RoboDK station: verify_station_copy.rdk

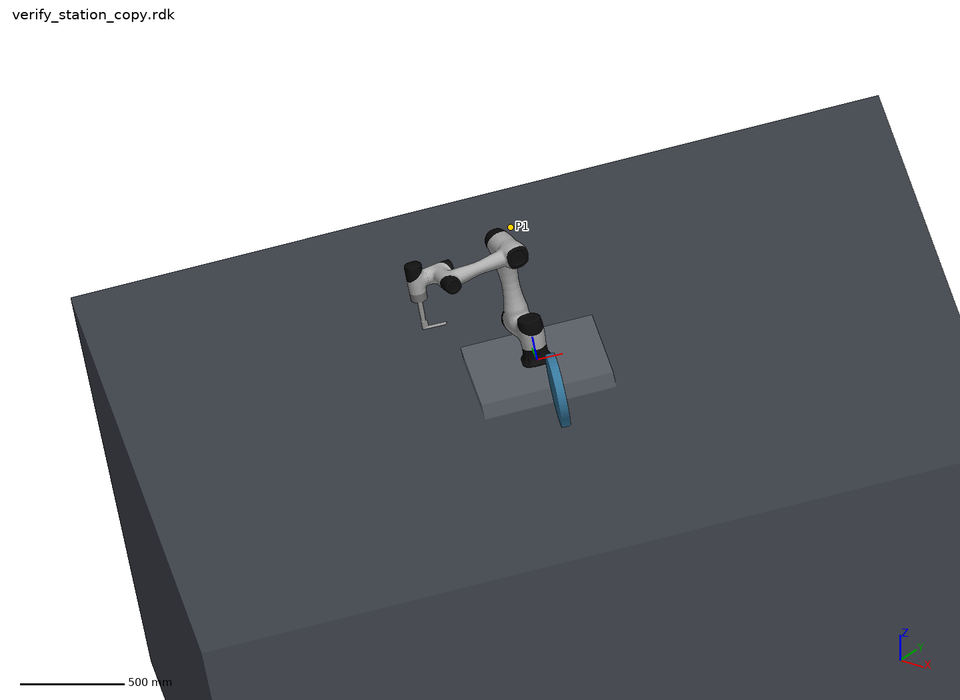
[picture v0: the station drawn from its stored meshes, robots at their saved joint values, targets as dots, program paths as lines]
Station 新建工作站 (1) (saved by RoboDK 5.9.0). Poses are relative to the parent item; angles as X-Y-Z fixed-axis rotations.
Station parameters (name, value as stored): Trace_Render_Style, 0
  - Python program TCP真实运动_升级前备份_20260910_170410 (listed below)
  - Python program 方向角计算 (listed below)
  - frame Dobot CR5 Base at (213.88, 904.45, 25.18) mm, rotated rx -0.42 ry -9.85 rz 44.17 deg
    - robot Dobot CR5: 6 axes, payload 5 kg, reach 900 mm, repeatability 0.03 mm, weight 23 kg
        modified DH rows (alpha deg, a mm, theta deg, d mm): 0, 0, 0, 147; 90, 0, 90, 0; 0, 427, 0, 0; 0, 357, -90, 141; -90, 0, 0, 116; 90, 0, 180, 100.5
        joint limits [-360, -360, -160, -360, -360, -360] to [360, 360, 160, 360, 360, 360]; home [0, 0, -90, 90, 90, 0]; saved at [-163.62, -0.936, -91.282, 2.218, 90, 106.38]
      - tool , TCP at (0, 0, 159.63) mm, size 120.1 x 159.6 x 24.6 mm, geometry from bs1.stp
    - target P1 (joint target) at (-20.1, -241.48, 846.75) mm, rotated rx -90 ry 1.35 rz 179.96 deg; joints [0, -37.451, 84.112, -46.661, 0, 0] of Dobot CR5
    - object  at (0, 0, 0) mm, rotated rx 0 ry -1.35 rz -0.05 deg, size 650 x 650 x 80 mm
    - object  at (0, 0, 0) mm, rotated rx 0 ry -1.35 rz -0.05 deg, size 4000 x 4000 x 2000 mm
    - object  at (0, -956, 300) mm, rotated rx 139.77 ry 89.72 rz -40.3 deg, size 360 x 360 x 40 mm
  - Python program TCP仿真_升级前备份_20260909_173616 (listed below)
  - Python program TCP仿真_升级前备份_20260910_161757 (listed below)
  - Python program TCP仿真_升级前备份_20260910_164419 (listed below)
  - Python program test (listed below)
  - Python program 机械臂法兰真实运动 (listed below)
  - Python program TCP真实运动_到位复核前备份_20260910_172919 (listed below)
  - Python program TCP真实运动 (listed below)
  - Python program TCP仿真_退让换向升级前 (listed below)
  - Python program TCP仿真 (listed below)
  - Python program 机械臂TCP仿真_副本 (listed below)

--- Python program TCP真实运动_升级前备份_20260910_170410 ---
# -*- coding: utf-8 -*-
"""
RoboDK 实机运动控制（基于 robodk_movej_diag.py 的成功模式）
- 单点：TCP 输入 -> IK 检测 -> MoveL/MoveJ 执行
- 连续轨迹：坐标列表 -> 逐点 IK 检测 -> MoveJ+MoveL 序列
模式：RUNMODE_RUN_ROBOT + robot.Connect()
"""

from robodk.robolink import *
from robodk.robomath import *
import tkinter as tk
from tkinter import ttk, scrolledtext, filedialog
import time
import math
import json

ROBOT_SPEED = 20.0
NL = chr(10)

RDK = Robolink()

def fanuc_to_pose(x, y, z, rx, ry, rz):
    return Fanuc_2_Pose([x, y, z, rx, ry, rz])

def pose_to_fanuc(pose):
    return Pose_2_Fanuc(pose)

# ---- 获取机器人 ----
robot = RDK.Item('', ITEM_TYPE_ROBOT)
if not robot.Valid():
    raise Exception("未找到机器人")

# ---- 全局变量 ----
text_points = None
text_log = None
record_text = None
entries_single = None
entries_joint = None
move_type = None
trajectory_records = []
_connected = False

# ============================================================
# 日志
# ============================================================
def log(s):
    print(s)
    if text_log:
        text_log.insert(tk.END, str(s) + NL)
        text_log.see(tk.END)
        root.update_idletasks()

# ============================================================
# 连接（只连一次，复用）
# ============================================================
def ensure_connected():
    global _connected
    if _connected:
        return True
    try:
        robot.Connect()
        time.sleep(1.5)
        status, msg = robot.ConnectedState()
        log("连接状态: %s, %s" % (status, msg))
        RDK.setRunMode(RUNMODE_RUN_ROBOT)
        log("RunMode: %s" % RDK.RunMode())
        if status < 0:
            _connected = False
            log("机器人连接未建立，状态=%s：%s" % (status, msg))
            return False
        _connected = True
        return True
    except Exception as e:
        log("连接失败: %s" % e)
        return False

# ============================================================
# 解析坐标
# ============================================================
def parse_points():
    if not text_points:
        return []
    raw = text_points.get("1.0", tk.END)
    points = []
    for line in raw.strip().split(NL):
        line = line.strip()
        if not line or line.startswith("#"):
            continue
        try:
            vals = [float(v.strip()) for v in line.split(",")]
            if len(vals) >= 6:
                points.append(vals[:6])
        except ValueError:
            pass
    return points

# ============================================================
# 读取当前位置
# ============================================================
def read_current(entries=None):
    try:
        pose = robot.Pose()
        v = pose_to_fanuc(pose)
        log("")
        log("当前 TCP：X=%.3f Y=%.3f Z=%.3f Rx=%.3f Ry=%.3f Rz=%.3f" % tuple(v[:6]))
    except Exception as e:
        log("读取失败：%s" % e)

def fill_current(entries=None):
    try:
        pose = robot.Pose()
        v = pose_to_fanuc(pose)
        if entries:
            for e, val in zip(entries, v):
                e.delete(0, tk.END)
                e.insert(0, "%.3f" % val)
        log("当前 TCP 已填入")
    except Exception as e:
        log("读取失败：%s" % e)

# ============================================================
# IK 检测
# 注意：SolveIK 显式使用当前 Tool + Reference，和 MoveL/MoveJ 保持一致。
# ============================================================
def check_ik_single(entries=None):
    if not entries:
        return
    try:
        values = [float(e.get()) for e in entries]
    except ValueError:
        log("输入无效")
        return

    x, y, z, rx, ry, rz = values
    target = fanuc_to_pose(x, y, z, rx, ry, rz)
    log("")
    log("目标：X=%.3f Y=%.3f Z=%.3f Rx=%.3f Ry=%.3f Rz=%.3f" % (x, y, z, rx, ry, rz))

    try:
        tool_pose = robot.PoseTool()
        frame_pose = robot.PoseFrame()
        joints = robot.SolveIK(target, tool=tool_pose, reference=frame_pose)
        if joints is None:
            log("IK 不可达")
        else:
            q = joints.list()
            if len(q) < 6:
                log("IK 返回关节数量异常：%d，原始数据=%r" % (len(q), q))
                return
            log("IK 可达")
            log("  关节：J1=%.2f J2=%.2f J3=%.2f J4=%.2f J5=%.2f J6=%.2f" % tuple(q[:6]))
    except Exception as e:
        log("检测失败：%s" % e)

def check_all_ik():
    points = parse_points()
    if not points:
        log("没有有效点")
        return

    log("")
    log("========== 检测全部 %d 个点 ==========" % len(points))
    all_ok = True
    for i, p in enumerate(points):
        try:
            target = fanuc_to_pose(*p)
            joints = robot.SolveIK(target, tool=robot.PoseTool(), reference=robot.PoseFrame())
            if joints is None:
                log("  P%d: 不可达" % (i+1))
                all_ok = False
            else:
                q = joints.list()
                if len(q) < 6:
                    raise ValueError("IK 返回关节数量异常: %d, raw=%r" % (len(q), q))
                log("  P%d: 可达  J1=%.1f J2=%.1f J3=%.1f J4=%.1f J5=%.1f J6=%.1f" % (i+1, *q[:6]))
        except Exception as e:
            log("  P%d: 检测失败 %s" % (i+1, e))
            all_ok = False
    if all_ok:
        log("全部 %d 个点可达" % len(points))
    else:
        log("存在不可达点，执行时会跳过")

# ============================================================
# 执行单点
# ============================================================
def execute_single(entries=None, mtype="MoveL"):
    if not entries:
        return
    try:
        values = [float(e.get()) for e in entries]
    except ValueError:
        log("输入无效")
        return

    x, y, z, rx, ry, rz = values
    target = fanuc_to_pose(x, y, z, rx, ry, rz)
    log("")
    log("目标：X=%.3f Y=%.3f Z=%.3f Rx=%.3f Ry=%.3f Rz=%.3f" % (x, y, z, rx, ry, rz))

    try:
        tool_pose = robot.PoseTool()
        frame_pose = robot.PoseFrame()
        joints = robot.SolveIK(target, tool=tool_pose, reference=frame_pose)
        if joints is None:
            log("IK 不可达，取消执行")
            return
        q = joints.list()
        if len(q) < 6:
            log("IK 返回关节数量异常：%d，取消执行；原始数据=%r" % (len(q), q))
            return
        log("IK 可达：J1=%.2f J2=%.2f J3=%.2f J4=%.2f J5=%.2f J6=%.2f" % tuple(q[:6]))
    except Exception as e:
        log("IK 检查失败：%s" % e)
        return

    if not ensure_connected():
        return

    try:
        robot.setPoseFrame(robot.PoseFrame())
        robot.setPoseTool(robot.PoseTool())
        robot.setSpeed(ROBOT_SPEED)
        log("发送 %s..." % mtype)
        if mtype == "MoveJ":
            robot.MoveJ(target)
        else:
            robot.MoveL(target)
        log("执行完成")
    except Exception as e:
        log("失败: %s: %s" % (type(e).__name__, e))

# ============================================================
# 连续运动：选项卡3直接输入 TCP / 关节点，逐点检查后加入轨迹
# ============================================================
trajectory_records = []
record_text = None
traj_entries = None
traj_type = None
singular_var = None
j6_direction_var = None


def _parse_six_from_entries(entries, label):
    if not entries or len(entries) != 6:
        log("%s输入框异常：需要 6 个值" % label)
        return None
    try:
        vals = [float(e.get().strip()) for e in entries]
    except (ValueError, AttributeError):
        log("%s输入无效：6 个值必须全部为数字" % label)
        return None
    if not all(math.isfinite(v) for v in vals):
        log("%s输入无效：不能包含 NaN 或无穷值" % label)
        return None
    return vals


def _check_tcp_reachable(vals):
    """检查单个 TCP 点 IK 是否可达，返回 (True, target, joints)。"""
    try:
        target = fanuc_to_pose(*vals)
        tool_pose = robot.PoseTool()
        frame_pose = robot.PoseFrame()
        joints = robot.SolveIK(target, tool=tool_pose, reference=frame_pose)

        if joints is None:
            log("TCP IK：不可达")
            return False, None, None

        q = joints.list()
        if len(q) < 6:
            log("TCP IK：返回关节数量异常：%r" % q)
            return False, None, None

        log("TCP IK：可达")
        log("  IK关节：J1=%.2f J2=%.2f J3=%.2f J4=%.2f J5=%.2f J6=%.2f" % tuple(q[:6]))
        return True, target, q[:6]
    except Exception as e:
        log("TCP IK 检查失败：%s: %s" % (type(e).__name__, e))
        return False, None, None


def _check_tcp_segment_continuous(prev_vals, curr_vals, segment_index, samples=20):
    """检查前一个 TCP 点到当前 TCP 点之间的整段插补路径 IK 连续可达性。

    暂不考虑障碍物，只对 TCP 位姿做线性插值，并对每个采样位姿执行 SolveIK。
    起点和终点也包含在采样检查中。
    """
    if prev_vals is None:
        return True

    log("开始检查 P%d -> P%d 的 TCP 连续 IK（%d 个采样点）" %
        (segment_index - 1, segment_index, samples + 1))

    tool_pose = robot.PoseTool()
    frame_pose = robot.PoseFrame()

    for k in range(samples + 1):
        t = float(k) / float(samples)
        vals = [prev_vals[i] + (curr_vals[i] - prev_vals[i]) * t for i in range(6)]
        try:
            pose = fanuc_to_pose(*vals)
            joints = robot.SolveIK(pose, tool=tool_pose, reference=frame_pose)
            if joints is None:
                log("  P%d -> P%d：第 %d/%d 个采样点 IK 不可达，t=%.3f" %
                    (segment_index - 1, segment_index, k + 1, samples + 1, t))
                log("  TCP：X=%.3f Y=%.3f Z=%.3f Rx=%.3f Ry=%.3f Rz=%.3f" % tuple(vals))
                return False
            q = joints.list()
            if len(q) < 6:
                log("  P%d -> P%d：第 %d 个采样点 IK 返回异常：%r" %
                    (segment_index - 1, segment_index, k + 1, q))
                return False
        except Exception as e:
            log("  P%d -> P%d：第 %d 个采样点 IK 检查失败：%s: %s" %
                (segment_index - 1, segment_index, k + 1, type(e).__name__, e))
            return False

    log("P%d -> P%d：连续 IK 检查通过" % (segment_index - 1, segment_index))
    return True


def _check_joint_reachable(q):
    """兼容旧代码：关节点不做可达性/限位检查，输入合法即可加入。"""
    return True


def refresh_record_list():
    if record_text is None:
        return

    record_text.delete("1.0", tk.END)

    for i, rec in enumerate(trajectory_records, 1):
        kind = rec["type"]
        vals = rec["values"]

        if kind == "TCP":
            mark = " [J6特异点 %s180°]" % ("+" if rec.get("j6_delta", 180) >= 0 else "-") if rec.get("singular", False) else ""
            record_text.insert(
                tk.END,
                "P%-3d [TCP]%s   X=%9.3f Y=%9.3f Z=%9.3f Rx=%8.3f Ry=%8.3f Rz=%8.3f%s" %
                (i, mark, *vals, NL)
            )
        else:
            record_text.insert(
                tk.END,
                "P%-3d [JNT]   J1=%8.3f J2=%8.3f J3=%8.3f J4=%8.3f J5=%8.3f J6=%8.3f%s" %
                (i, *vals, NL)
            )


def add_and_check_trajectory_point():
    """
    选项卡3逐点输入：
    - 普通 TCP：立即做端点 IK，并检查与前一个普通 TCP 点之间的连续 IK。
    - TCP 末端特异点：跳过 IK；要求与前一个普通 TCP 点 XYZ 相同，执行时仅 J6 转 ±180°。
    - 关节：不做 IK/限位检查，只将角度规范到 (-180°, 180°]。
    注意：这些检查只在“加入点”时完成；正式实机执行时不再做轨迹预检。
    """
    kind = traj_type.get()
    vals = _parse_six_from_entries(traj_entries, kind)
    if vals is None:
        return

    log("")
    log("========== 检查连续运动第 %d 点 ==========" % (len(trajectory_records) + 1))

    is_singular = bool(singular_var.get()) if (kind == "TCP" and singular_var is not None) else False
    j6_delta = int(j6_direction_var.get()) if (j6_direction_var is not None) else 180

    if kind == "TCP" and is_singular:
        if not trajectory_records:
            log("末端特异点不能作为第一个点：需要先有一个起始运动点。")
            return
        prev = trajectory_records[-1]
        if prev["type"] != "TCP" or prev.get("singular", False):
            log("末端特异点前一项必须是普通 TCP 点。")
            return
        prev_vals = prev["values"]
        pos_err = math.sqrt(sum((vals[k] - prev_vals[k]) ** 2 for k in range(3)))
        if pos_err > 1e-3:
            log("末端特异点未加入：XYZ 必须与前一个普通 TCP 点相同。")
            log("  与前一点位置差：%.6f mm" % pos_err)
            return
        try:
            target = fanuc_to_pose(*vals)
        except Exception as e:
            log("末端特异点姿态转换失败：%s: %s" % (type(e).__name__, e))
            return

        trajectory_records.append({
            "type": "TCP", "values": vals[:], "target": target, "joints": None,
            "singular": True, "j6_delta": j6_delta,
        })
        log("P%d [TCP-特异点]：已加入，跳过 IK。" % len(trajectory_records))
        log("  执行时保持 J1~J5 不变，仅让 J6 转 %+d°。" % j6_delta)
        if singular_var is not None:
            singular_var.set(False)
        refresh_record_list()
        return

    if kind == "TCP":
        ok, target, joints = _check_tcp_reachable(vals)
        if not ok:
            log("该 TCP 点未加入轨迹。")
            return

        # 只在点加入阶段检查连续 IK；实机正式执行时不再重复预检。
        if trajectory_records and trajectory_records[-1]["type"] == "TCP" and not trajectory_records[-1].get("singular", False):
            prev_vals = trajectory_records[-1]["values"]
            segment_no = len(trajectory_records) + 1
            if not _check_tcp_segment_continuous(prev_vals, vals, segment_no, samples=20):
                log("P%d [TCP]：上一普通 TCP 点到当前点的连续 IK 检查失败，该点未加入轨迹。" % segment_no)
                return

        trajectory_records.append({
            "type": "TCP", "values": vals[:], "target": target, "joints": joints,
            "singular": False, "j6_delta": 0,
        })
        log("P%d [TCP]：检查通过，已加入连续运动。" % len(trajectory_records))
    else:
        corrected = []
        for v in vals:
            v = ((v + 180.0) % 360.0) - 180.0
            if v <= -180.0:
                v = 180.0
            corrected.append(v)
        if corrected != vals:
            log("关节点角度已自动纠正到 (-180°, 180°]：")
            log("  原始：" + "  ".join("J%d=%+.3f°" % (i + 1, vals[i]) for i in range(6)))
            log("  修正：" + "  ".join("J%d=%+.3f°" % (i + 1, corrected[i]) for i in range(6)))
        trajectory_records.append({
            "type": "JOINT", "values": corrected[:], "target": None, "joints": corrected[:],
            "singular": False, "j6_delta": 0,
        })
        log("P%d [JNT]：未做 IK 检查，角度规范化后已加入连续运动。" % len(trajectory_records))

    refresh_record_list()


def _write_values_to_traj_entries(values, label):
    if not traj_entries or len(traj_entries) != 6:
        log("连续运动输入框异常：无法写入当前%s" % label)
        return False
    for e, val in zip(traj_entries, values[:6]):
        e.delete(0, tk.END)
        e.insert(0, "%.3f" % float(val))
    log("当前%s已写入选项卡3输入框" % label)
    return True


def read_current_tcp_to_traj():
    """读取当前 RoboDK TCP，并写入选项卡3的 TCP 输入框。"""
    try:
        pose = robot.Pose()
        vals = pose_to_fanuc(pose)
        log("========== 读取当前 TCP -> 选项卡3 ==========")
        log("X=%+.3f Y=%+.3f Z=%+.3f Rx=%+.3f Ry=%+.3f Rz=%+.3f" % tuple(vals))
        if traj_type.get() != "TCP":
            traj_type.set("TCP")
            _update_traj_labels_and_defaults()
        return _write_values_to_traj_entries(vals, "TCP")
    except Exception as e:
        log("读取当前 TCP 失败：%s: %s" % (type(e).__name__, e))
        return False


def read_current_joints_to_traj():
    """读取 RoboDK Robot Item 当前关节，并写入选项卡3的关节输入框。"""
    q = read_current_joints(None)
    if q is None or len(q) < 6:
        return False
    log("========== 读取当前关节 -> 选项卡3 ==========")
    if traj_type.get() != "JOINT":
        traj_type.set("JOINT")
        _update_traj_labels_and_defaults()
    return _write_values_to_traj_entries(q, "关节")


def clear_trajectory_input():
    if not traj_entries:
        return

    for e in traj_entries:
        e.delete(0, tk.END)

    if traj_type.get() == "TCP":
        defaults = ["0.000", "-241.500", "1047.000", "-90.000", "0.000", "180.000"]
    else:
        defaults = ["0.000"] * 6

    for e, val in zip(traj_entries, defaults):
        e.insert(0, val)




def import_trajectory():
    """
    从仿真程序导出的 JSON 轨迹文件导入到实机连续运动列表。

    重要：这里不做连续轨迹预检，不做 MoveJ TCP 轨迹预检。
    普通 TCP 如果 JSON 中没有保存 IK 关节，则只针对该点单独 SolveIK，
    用于得到实机执行所需的目标关节；这不是连续轨迹预检。
    """
    filepath = filedialog.askopenfilename(
        title="导入仿真轨迹",
        defaultextension=".json",
        filetypes=[("JSON 轨迹文件", "*.json"), ("所有文件", "*.*")]
    )
    if not filepath:
        return

    try:
        with open(filepath, "r", encoding="utf-8") as f:
            data = json.load(f)

        if not isinstance(data, list):
            raise ValueError("轨迹文件顶层必须是列表。")

        imported = []
        for idx, item in enumerate(data, 1):
            if not isinstance(item, dict):
                raise ValueError("P%d 不是对象格式。" % idx)

            kind = str(item.get("type", "")).upper()
            if kind == "JNT":
                kind = "JOINT"
            if kind not in ("TCP", "JOINT"):
                raise ValueError("P%d type 不支持：%r" % (idx, item.get("type")))

            values = item.get("values")
            if not isinstance(values, list) or len(values) != 6:
                raise ValueError("P%d values 必须是长度为6的列表。" % idx)
            try:
                values = [float(v) for v in values]
            except (TypeError, ValueError):
                raise ValueError("P%d values 必须全部为数字。" % idx)
            if not all(math.isfinite(v) for v in values):
                raise ValueError("P%d values 不能包含 NaN 或无穷值。" % idx)

            is_singular = bool(item.get("singular", False)) and kind == "TCP"
            j6_delta = int(item.get("j6_delta", 180)) if is_singular else 0
            if is_singular and j6_delta not in (-180, 180):
                raise ValueError("P%d 特异点 j6_delta 只能是 +180 或 -180。" % idx)

            if kind == "JOINT":
                # 与手动输入保持一致：自动规范到 (-180,180]。
                corrected = []
                for v in values:
                    v = ((v + 180.0) % 360.0) - 180.0
                    if v <= -180.0:
                        v = 180.0
                    corrected.append(v)
                values = corrected
                imported.append({
                    "type": "JOINT", "values": values, "target": None,
                    "joints": values[:], "singular": False, "j6_delta": 0
                })
                continue

            target = fanuc_to_pose(*values)

            if is_singular:
                # 特异点严格要求前一项为普通 TCP，且 XYZ 相同。
                if not imported:
                    raise ValueError("P%d 末端特异点不能作为第一个点。" % idx)
                prev = imported[-1]
                if prev["type"] != "TCP" or prev.get("singular", False):
                    raise ValueError("P%d 末端特异点前一项必须是普通 TCP。" % idx)
                pos_err = math.sqrt(sum((values[k] - prev["values"][k]) ** 2 for k in range(3)))
                if pos_err > 1e-3:
                    raise ValueError("P%d 末端特异点 XYZ 必须与前一个普通 TCP 相同，位置差 %.6f mm。" % (idx, pos_err))
                imported.append({
                    "type": "TCP", "values": values[:], "target": target,
                    "joints": None, "singular": True, "j6_delta": j6_delta
                })
                continue

            # 优先使用文件中可能保存的 IK；当前仿真脚本的 JSON 通常没有 joints，
            # 因此回退到“单点 SolveIK”，仅为了得到实机 MoveJ/MoveL 所需目标关节。
            q = item.get("joints")
            if isinstance(q, list) and len(q) >= 6:
                try:
                    q = [float(v) for v in q[:6]]
                    if not all(math.isfinite(v) for v in q):
                        q = None
                except (TypeError, ValueError):
                    q = None

            if q is None:
                joints = robot.SolveIK(
                    target, tool=robot.PoseTool(), reference=robot.PoseFrame()
                )
                if joints is None:
                    raise ValueError("P%d 普通 TCP 单点 IK 无解，无法导入。" % idx)
                q = joints.list()
                if q is None or len(q) < 6:
                    raise ValueError("P%d 普通 TCP IK 返回关节数量异常：%r" % (idx, q))
                q = [float(v) for v in q[:6]]

            imported.append({
                "type": "TCP", "values": values[:], "target": target,
                "joints": q[:], "singular": False, "j6_delta": 0
            })

        trajectory_records.clear()
        trajectory_records.extend(imported)
        refresh_record_list()
        log("")
        log("========== 导入仿真轨迹 ==========")
        log("文件：%s" % filepath)
        log("已导入 %d 个轨迹点。" % len(imported))
        log("连续轨迹预检：未执行（按实机程序设计）。")
        log("普通 TCP：仅在缺少保存IK时进行单点 SolveIK；不进行连续段预检。")
        log("末端特异点：跳过IK，仅保留 J6 ±180° 标记。")
        log("================================")
    except Exception as e:
        log("轨迹导入失败：%s: %s" % (type(e).__name__, e))

def delete_last_record():
    if trajectory_records:
        rec = trajectory_records.pop()
        refresh_record_list()
        log("已删除最后一点：P%d [%s]" %
            (len(trajectory_records) + 1, rec["type"]))
    else:
        log("当前没有可删除的连续运动点")


def clear_records():
    trajectory_records.clear()
    refresh_record_list()
    log("连续运动点列表已清空")


def execute_recorded_trajectory():
    """
    实机执行选项卡3轨迹。

    重要：不做仿真轨迹预检。TCP 的 IK/连续 IK 已在“检查并加入当前点”阶段完成，
    实机这里只负责按仿真已经验证过的顺序执行。

    普通 TCP：第一个 TCP MoveJ，后续普通 TCP 优先 MoveL；MoveL 失败后直接用已经保存的 IK 关节 MoveJ 兜底。
    末端特异点：跳过 IK，读取当前 RoboDK Robot Item 关节，仅 J6 转 ±180°。
    特异点后的普通 TCP：重新使用该普通 TCP 自己保存的 IK，正常 MoveL。
    关节点：直接 MoveJ。
    StoppedError: Robot not connected：继续视为本段结束标志。
    """
    if not trajectory_records:
        log("没有已检查通过的运动点，请先在选项卡3输入并加入点。")
        return

    log("")
    log("========== 执行实机连续运动：%d 个点 ==========" % len(trajectory_records))
    log("轨迹预检：跳过（已在仿真/加入点阶段完成）")

    if not ensure_connected():
        log("连续运动取消：机器人未连接")
        return

    try:
        RDK.setRunMode(RUNMODE_RUN_ROBOT)
        robot.setPoseFrame(robot.PoseFrame())
        robot.setPoseTool(robot.PoseTool())
        robot.setSpeed(ROBOT_SPEED)

        tcp_count = 0
        completed_count = 0

        for i, rec in enumerate(trajectory_records, 1):
            kind = rec["type"]
            vals = rec["values"]
            is_singular = bool(rec.get("singular", False))
            j6_delta = int(rec.get("j6_delta", 180))

            if kind == "TCP" and is_singular:
                move_name = "J6特异点"
            elif kind == "TCP":
                move_name = "MoveJ" if tcp_count == 0 else "MoveL"
            else:
                move_name = "MoveJ"

            log("")
            log("---- 开始执行 P%d [%s] -> %s ----" % (i, kind, move_name))

            try:
                if kind == "TCP":
                    if is_singular:
                        # 特异点：当前 RoboDK Robot Item 关节作为起点，保持 J1~J5，仅改变 J6。
                        current_q = list(robot.SimulatorJoints())
                        if len(current_q) < 6:
                            raise RuntimeError("特异点：RoboDK SimulatorJoints 返回关节数量不足6个：%r" % current_q)
                        current_q = current_q[:6]
                        q_special = current_q[:]
                        q_special[5] += float(j6_delta)
                        # 保持与前面关节点规范一致，避免无意义多圈累加。
                        q_special[5] = ((q_special[5] + 180.0) % 360.0) - 180.0
                        if q_special[5] <= -180.0:
                            q_special[5] = 180.0
                        log("P%d [TCP-特异点]：J6 %.3f° -> %.3f°，J1~J5保持不变" %
                            (i, current_q[5], q_special[5]))
                        robot.MoveJ(q_special)
                        tcp_count += 1
                    elif tcp_count == 0:
                        # 首个普通TCP：使用加入阶段已经得到的IK关节，避免再次SolveIK。
                        q = rec.get("joints")
                        if q is None or len(q) < 6:
                            raise RuntimeError("P%d：缺少已保存的 TCP IK 关节解。" % i)
                        robot.MoveJ(q[:6])
                        tcp_count += 1
                    else:
                        # 后续普通TCP：优先 MoveL。
                        target = rec.get("target")
                        q = rec.get("joints")
                        if target is None or q is None or len(q) < 6:
                            raise RuntimeError("P%d：缺少已保存的 TCP 目标位姿或 IK 关节解。" % i)
                        try:
                            robot.MoveL(target)
                        except Exception as e_l:
                            # 仿真已经检查过 MoveJ 的 TCP 轨迹，因此实机不再重复预检，直接用已验证的 IK 解兜底。
                            log("P%d [TCP] -> MoveL 失败：%s: %s" % (i, type(e_l).__name__, e_l))
                            log("P%d [TCP] -> 直接使用仿真已验证的 IK 关节解执行 MoveJ 兜底。" % i)
                            robot.MoveJ(q[:6])

                else:
                    q = rec["values"][:6]
                    robot.MoveJ(q)

                completed_count += 1
                log("P%d [%s] -> %s 返回正常，进入下一段。" % (i, kind, move_name))

            except Exception as e:
                err_type = type(e).__name__
                err_text = str(e)
                if err_type == "StoppedError" and "Robot not connected" in err_text:
                    completed_count += 1
                    log("P%d [%s] -> %s 已结束。" % (i, kind, move_name))
                    log("收到结束标志：StoppedError: Robot not connected")
                    log("将该报错视为本段运动结束，继续执行下一段。")
                    continue

                log("P%d [%s] -> %s 执行失败：%s: %s" %
                    (i, kind, move_name, err_type, err_text))
                log("非预期错误，停止后续连续运动。")
                return

        log("")
        log("========== 实机连续运动执行完成：%d/%d 段 ==========" %
            (completed_count, len(trajectory_records)))

    except Exception as e:
        log("连续运动初始化失败：%s: %s" % (type(e).__name__, e))


# 保留旧函数名，避免其他代码调用失效。
def execute_trajectory():
    execute_recorded_trajectory()


# ============================================================
# 实机关节运动
# ============================================================
def _joint_values_from_entries(entries):
    """从 GUI 读取 J1~J6 目标角度。单位：deg。"""
    if not entries or len(entries) != 6:
        log("目标关节输入框异常：需要 J1~J6 共 6 个")
        return None
    try:
        q = [float(e.get().strip()) for e in entries]
    except (ValueError, AttributeError):
        log("目标关节输入无效：J1~J6 必须全部填写数字")
        return None
    if not all(math.isfinite(v) for v in q):
        log("目标关节输入无效：不能包含 NaN 或无穷值")
        return None
    return q


def read_current_joints(entries=None):
    """读取 RoboDK Robot Item 当前关节值，并可直接填入 J1~J6 输入框。
    注意：这里读取的是 RoboDK 当前 Robot Item 的关节状态，不调用 CR5 控制器 GetAngle。
    """
    try:
        joints = robot.SimulatorJoints()
        q = list(joints) if hasattr(joints, "__iter__") else [joints]
        if len(q) < 6:
            log("读取当前关节失败：SimulatorJoints 返回 %r" % (q,))
            log("请确认 RoboDK 窗口中的机器人已经连接并显示实时关节角度。")
            return None

        q = q[:6]
        log("")
        log("========== RoboDK 当前关节 ==========")
        log("J1=%+.3f°  J2=%+.3f°  J3=%+.3f°" % tuple(q[:3]))
        log("J4=%+.3f°  J5=%+.3f°  J6=%+.3f°" % tuple(q[3:]))

        if entries and len(entries) == 6:
            for e, val in zip(entries, q):
                e.delete(0, tk.END)
                e.insert(0, "%.3f" % val)
            log("当前关节已填入 J1~J6 输入框")

        return q
    except Exception as e:
        log("读取 RoboDK 当前关节失败：%s: %s" % (type(e).__name__, e))
        return None


def fill_current_joints(entries=None):
    """当前 RoboDK 关节 -> 目标关节输入框。"""
    return read_current_joints(entries)


def execute_joint_target(entries=None):
    """按 GUI 输入的 J1~J6 目标角度直接执行实机 MoveJ，不经过 TCP/IK。"""
    q = _joint_values_from_entries(entries)
    if q is None:
        return

    log("")
    log("========================================")
    log("====== 实机指定关节角度 MoveJ ======")
    log("目标：J1=%+.3f°  J2=%+.3f°  J3=%+.3f°" % tuple(q[:3]))
    log("      J4=%+.3f°  J5=%+.3f°  J6=%+.3f°" % tuple(q[3:]))
    log("运动速度：%.1f" % ROBOT_SPEED)
    log("控制方式：RoboDK Robot Item -> RUNMODE_RUN_ROBOT -> MoveJ(q)")

    if not ensure_connected():
        log("实机关节运动取消：机器人未连接")
        return

    try:
        RDK.setRunMode(RUNMODE_RUN_ROBOT)
        log("RunMode：%s" % RDK.RunMode())
        robot.setSpeed(ROBOT_SPEED)
        log("发送 MoveJ 目标：%r" % q)
        robot.MoveJ(q)
        log("MoveJ 命令已发送，目标关节角度：%r" % q)
        log("========================================")
    except Exception as e:
        log("实机 MoveJ 失败：%s: %s" % (type(e).__name__, e))


def clear_joint_target(entries=None):
    if not entries:
        return
    for e in entries:
        e.delete(0, tk.END)
        e.insert(0, "0.000")
    log("目标关节输入已清零")

# ============================================================
# GUI
# ============================================================
root = tk.Tk()
root.title("RoboDK - 机械臂运动控制")
root.geometry("1200x750")
root.resizable(True, True)

tk.Label(root, text="Dobot CR5 运动控制", font=("Microsoft YaHei", 16, "bold")).pack(pady=10)

notebook = ttk.Notebook(root)
notebook.pack(fill=tk.BOTH, expand=True, padx=10, pady=5)

# ---- 选项卡 1：单点运动 ----
tab_single = ttk.Frame(notebook)
notebook.add(tab_single, text="单点运动")

frame_coord = tk.LabelFrame(tab_single, text="目标 TCP（Fanuc 格式）")
frame_coord.pack(fill=tk.X, padx=10, pady=10)

names = ["X (mm)", "Y (mm)", "Z (mm)", "Rx (deg)", "Ry (deg)", "Rz (deg)"]
defaults = ["0.000", "-241.500", "1047.000", "-90.000", "0.000", "180.000"]
entries_single = []

for i in range(6):
    tk.Label(frame_coord, text=names[i]).grid(row=0, column=i*2, padx=5, pady=10)
    e = tk.Entry(frame_coord, width=12)
    e.insert(0, defaults[i])
    e.grid(row=0, column=i*2+1, padx=5, pady=10)
    entries_single.append(e)

frame_mtype = tk.Frame(tab_single)
frame_mtype.pack(fill=tk.X, padx=10, pady=5)
move_type = tk.StringVar(value="MoveL")
tk.Radiobutton(frame_mtype, text="MoveL (直线)", variable=move_type, value="MoveL").pack(side=tk.LEFT, padx=10)
tk.Radiobutton(frame_mtype, text="MoveJ (关节)", variable=move_type, value="MoveJ").pack(side=tk.LEFT, padx=10)

btn_single_frame = tk.Frame(tab_single)
btn_single_frame.pack(fill=tk.X, padx=10, pady=5)

def _read_current():
    read_current(entries_single)
def _fill_current():
    fill_current(entries_single)
def _check_ik():
    check_ik_single(entries_single)
def _exec_single():
    execute_single(entries_single, move_type.get())

tk.Button(btn_single_frame, text="读取当前 TCP", command=_read_current, width=15).pack(side=tk.LEFT, padx=3)
tk.Button(btn_single_frame, text="当前 TCP -> 输入框", command=_fill_current, width=20).pack(side=tk.LEFT, padx=3)
tk.Button(btn_single_frame, text="检测可达性", command=_check_ik, width=15, bg="#2196F3", fg="white").pack(side=tk.LEFT, padx=3)
tk.Button(btn_single_frame, text="执行运动", command=_exec_single, width=20,
          font=("Microsoft YaHei", 10, "bold"), bg="#4CAF50", fg="white").pack(side=tk.LEFT, padx=3)


# ---- 选项卡 2：目标关节运动（实机） ----
tab_joint = ttk.Frame(notebook)
notebook.add(tab_joint, text="目标关节运动")

frame_joint = tk.LabelFrame(tab_joint, text="目标关节（deg）")
frame_joint.pack(fill=tk.X, padx=10, pady=10)

joint_names = ["J1 (deg)", "J2 (deg)", "J3 (deg)", "J4 (deg)", "J5 (deg)", "J6 (deg)"]
joint_defaults = ["0.000", "0.000", "0.000", "0.000", "0.000", "0.000"]
entries_joint = []

for i in range(6):
    tk.Label(frame_joint, text=joint_names[i]).grid(row=0, column=i*2, padx=5, pady=10)
    e = tk.Entry(frame_joint, width=12)
    e.insert(0, joint_defaults[i])
    e.grid(row=0, column=i*2+1, padx=5, pady=10)
    entries_joint.append(e)

btn_joint_frame = tk.Frame(tab_joint)
btn_joint_frame.pack(fill=tk.X, padx=10, pady=8)

def _read_current_joint_values():
    read_current_joints(entries_joint)

def _fill_current_joints():
    fill_current_joints(entries_joint)

def _exec_joint():
    execute_joint_target(entries_joint)

def _zero_joints():
    clear_joint_target(entries_joint)

tk.Button(btn_joint_frame, text="读取当前关节", command=_read_current_joint_values, width=14).pack(side=tk.LEFT, padx=3)
tk.Button(btn_joint_frame, text="当前关节 -> 输入框", command=_fill_current_joints, width=20).pack(side=tk.LEFT, padx=3)
tk.Button(btn_joint_frame, text="执行指定关节 MoveJ", command=_exec_joint, width=24,
          font=("Microsoft YaHei", 10, "bold"), bg="#FF9800", fg="white").pack(side=tk.LEFT, padx=3)
tk.Button(btn_joint_frame, text="清零", command=_zero_joints, width=10).pack(side=tk.LEFT, padx=3)

tk.Label(tab_joint,
         text="输入 J1~J6 目标角度（deg），点击“执行指定关节 MoveJ”直接控制实机；不经过 TCP、Fanuc 转换或 IK。",
         fg="#555555").pack(anchor=tk.W, padx=15, pady=5)
tk.Label(tab_joint,
         text="安全提示：首次测试建议只改变一个关节、改变 5~10°，确认方向和角度定义正确后再进行大角度运动。",
         fg="#C62828").pack(anchor=tk.W, padx=15, pady=2)

# ---- 选项卡 3：连续运动 ----
tab_traj = ttk.Frame(notebook)
notebook.add(tab_traj, text="连续运动")

frame_traj_input = tk.LabelFrame(
    tab_traj,
    text="连续运动点输入：每次输入 1 个 TCP 点或 1 组关节角度，点击“检查并加入”"
)
frame_traj_input.pack(fill=tk.X, padx=10, pady=10)

type_frame = tk.Frame(frame_traj_input)
type_frame.pack(fill=tk.X, padx=8, pady=5)

tk.Label(type_frame, text="点类型：").pack(side=tk.LEFT, padx=3)

traj_type = tk.StringVar(value="TCP")
tk.Radiobutton(
    type_frame, text="TCP（X,Y,Z,Rx,Ry,Rz）",
    variable=traj_type, value="TCP"
).pack(side=tk.LEFT, padx=8)

tk.Radiobutton(
    type_frame, text="关节（J1~J6）",
    variable=traj_type, value="JOINT"
).pack(side=tk.LEFT, padx=8)

traj_names_tcp = ["X", "Y", "Z", "Rx", "Ry", "Rz"]
traj_names_joint = ["J1", "J2", "J3", "J4", "J5", "J6"]

traj_entries = []

# ---- 末端特异点设置 ----
singular_var = tk.BooleanVar(value=False)
j6_direction_var = tk.IntVar(value=180)

singular_frame = tk.Frame(frame_traj_input)
singular_frame.pack(fill=tk.X, padx=8, pady=3)

tk.Checkbutton(
    singular_frame,
    text="末端特异点（跳过IK，仅J6转180°）",
    variable=singular_var
).pack(side=tk.LEFT, padx=3)

tk.Label(singular_frame, text="J6方向：").pack(side=tk.LEFT, padx=(15, 3))
tk.Radiobutton(singular_frame, text="+180°", variable=j6_direction_var, value=180).pack(side=tk.LEFT, padx=3)
tk.Radiobutton(singular_frame, text="-180°", variable=j6_direction_var, value=-180).pack(side=tk.LEFT, padx=3)

# 输入框单独放在 grid 子容器中。
# frame_traj_input 本身使用 pack 管理子控件，不能再直接对它的子控件使用 grid。
traj_value_frame = tk.Frame(frame_traj_input)
traj_value_frame.pack(fill=tk.X, padx=8, pady=5)

for i in range(6):
    tk.Label(
        traj_value_frame,
        text=traj_names_tcp[i]
    ).grid(row=0, column=i * 2, padx=3, pady=8)

    e = tk.Entry(traj_value_frame, width=12)
    e.grid(row=0, column=i * 2 + 1, padx=4, pady=8)
    traj_entries.append(e)

# 默认先按 TCP 输入显示
tcp_defaults = ["0.000", "-241.500", "1047.000", "-90.000", "0.000", "180.000"]
for e, val in zip(traj_entries, tcp_defaults):
    e.insert(0, val)


def _update_traj_labels_and_defaults():
    """切换 TCP/关节输入时，更新标签和默认值。"""
    names = traj_names_tcp if traj_type.get() == "TCP" else traj_names_joint
    defaults = (
        tcp_defaults
        if traj_type.get() == "TCP"
        else ["0.000"] * 6
    )

    for i, e in enumerate(traj_entries):
        # grid 上的 Label 位于当前列
        for widget in traj_value_frame.grid_slaves(row=0, column=i * 2):
            widget.configure(text=names[i])

        e.delete(0, tk.END)
        e.insert(0, defaults[i])


tk.Radiobutton(
    type_frame, text="TCP（X,Y,Z,Rx,Ry,Rz）",
    variable=traj_type, value="TCP",
    command=_update_traj_labels_and_defaults
).pack_forget()

# 重新建立带 command 的两个单选按钮
for widget in list(type_frame.pack_slaves()):
    if isinstance(widget, tk.Radiobutton):
        widget.destroy()

tk.Radiobutton(
    type_frame, text="TCP（X,Y,Z,Rx,Ry,Rz）",
    variable=traj_type, value="TCP",
    command=_update_traj_labels_and_defaults
).pack(side=tk.LEFT, padx=8)

tk.Radiobutton(
    type_frame, text="关节（J1~J6）",
    variable=traj_type, value="JOINT",
    command=_update_traj_labels_and_defaults
).pack(side=tk.LEFT, padx=8)

btn_traj_input = tk.Frame(tab_traj)
btn_traj_input.pack(fill=tk.X, padx=10, pady=3)

tk.Button(
    btn_traj_input,
    text="检查并加入当前点",
    command=add_and_check_trajectory_point,
    width=22,
    bg="#2196F3",
    fg="white",
    font=("Microsoft YaHei", 10, "bold")
).pack(side=tk.LEFT, padx=3)

tk.Button(
    btn_traj_input,
    text="读取当前TCP并写入",
    command=read_current_tcp_to_traj,
    width=20
).pack(side=tk.LEFT, padx=3)

tk.Button(
    btn_traj_input,
    text="读取当前关节并写入",
    command=read_current_joints_to_traj,
    width=20
).pack(side=tk.LEFT, padx=3)

tk.Button(
    btn_traj_input,
    text="清空当前输入",
    command=clear_trajectory_input,
    width=16
).pack(side=tk.LEFT, padx=3)

tk.Label(
    tab_traj,
    text="输入一个点后：TCP 用 IK 判断可达；关节点不做检查，输入合法后直接加入。只有 TCP 检查通过的点或合法关节点才会加入下面列表。",
    fg="#555555"
).pack(anchor=tk.W, padx=15, pady=3)

frame_record = tk.LabelFrame(
    tab_traj,
    text="已检查通过的连续运动点（按加入顺序执行，可混合 TCP / 关节点）"
)
frame_record.pack(fill=tk.BOTH, expand=True, padx=10, pady=8)

record_text = tk.Text(frame_record, font=("Consolas", 10), height=10)
record_text.pack(fill=tk.BOTH, expand=True, padx=5, pady=5)

btn_record_frame = tk.Frame(tab_traj)
btn_record_frame.pack(fill=tk.X, padx=10, pady=4)

tk.Button(
    btn_record_frame, text="删除最后一点",
    command=delete_last_record, width=15
).pack(side=tk.LEFT, padx=3)

tk.Button(
    btn_record_frame, text="清空全部点",
    command=clear_records, width=15
).pack(side=tk.LEFT, padx=3)

tk.Button(
    btn_record_frame, text="导入轨迹",
    command=import_trajectory, width=14
).pack(side=tk.LEFT, padx=3)

tk.Button(
    btn_record_frame, text="执行整段连续运动",
    command=execute_recorded_trajectory,
    width=24,
    font=("Microsoft YaHei", 10, "bold"),
    bg="#4CAF50", fg="white"
).pack(side=tk.LEFT, padx=3)

tk.Label(
    tab_traj,
    text="执行：普通 TCP 首点 MoveJ、后续优先 MoveL；MoveL 失败直接用仿真已验证的 IK 解 MoveJ 兜底；末端特异点仅 J6 ±180°；关节点直接 MoveJ。实机不重复做轨迹预检。",
    fg="#555555"
).pack(anchor=tk.W, padx=15, pady=4)

# ---- 日志区 ----
frame_log = tk.LabelFrame(root, text="日志")
frame_log.pack(fill=tk.BOTH, expand=True, padx=10, pady=5)

text_log = scrolledtext.ScrolledText(frame_log, font=("Consolas", 10), height=8)
text_log.pack(fill=tk.BOTH, expand=True, padx=5, pady=5)

# ============================================================
# 启动
# ============================================================
log("机器人: " + robot.Name())
log("程序就绪。模式：RUNMODE_RUN_ROBOT + robot.Connect()")
log("单点：输入坐标 -> 检测可达性 -> 执行 MoveL/MoveJ")
log("目标关节：输入 J1~J6 -> 实机 MoveJ（不经过 TCP/Fanuc 转换和 IK）")
log("连续运动：支持导入仿真JSON；普通TCP使用仿真已验证IK（缺少时仅做单点SolveIK）；末端特异点跳过IK仅J6±180°；实机执行不重复轨迹预检；MoveL失败直接用仿真已验证IK解MoveJ兜底")

root.mainloop()

--- Python program 方向角计算 ---
import math
import tkinter as tk
from tkinter import ttk, messagebox

from robodk.robomath import Mat, Pose_2_Fanuc


# ============================================================
# 法兰坐标系 X+/Y+/Z+ -> RoboDK Fanuc/Motoman Rxyz
#
# 重要定义：
#   本程序现在不再只使用“末端朝向 Z 轴”计算姿态。
#   因为仅指定 Z+ 只能确定法兰朝向，不能确定绕 Z+ 的旋转。
#
#   现在可以同时输入：
#       X+ 在世界坐标中的方向
#       Y+ 在世界坐标中的方向
#       Z+ 在世界坐标中的方向
#
#   三个轴共同决定完整的法兰姿态。
#
#   如果只知道 Z+：
#       可以使用“Z+ + X+参考方向”模式，
#       程序会自动把 X+参考方向投影到垂直于 Z+ 的平面。
#
# 输出：
#   RoboDK Fanuc/Motoman [X,Y,Z,Rx,Ry,Rz]
#
# 单位：
#   输入向量：无单位，只表示方向
#   Rxyz：deg
# ============================================================


def vec_length(v):
    return math.sqrt(
        v[0] * v[0] +
        v[1] * v[1] +
        v[2] * v[2]
    )


def normalize(v):
    length = vec_length(v)

    if length < 1e-12:
        raise ValueError("方向向量不能为零向量")

    return (
        v[0] / length,
        v[1] / length,
        v[2] / length
    )


def dot(a, b):
    return (
        a[0] * b[0] +
        a[1] * b[1] +
        a[2] * b[2]
    )


def cross(a, b):
    return (
        a[1] * b[2] - a[2] * b[1],
        a[2] * b[0] - a[0] * b[2],
        a[0] * b[1] - a[1] * b[0]
    )


def scale(v, s):
    return (
        v[0] * s,
        v[1] * s,
        v[2] * s
    )


def sub(a, b):
    return (
        a[0] - b[0],
        a[1] - b[1],
        a[2] - b[2]
    )


def axis_to_rxyz(x_axis, y_axis, z_axis):
    """
    已知完整的法兰坐标系 X+/Y+/Z+ 在世界坐标中的方向，
    构造旋转矩阵并转换为 RoboDK Fanuc/Motoman Rxyz。
    """

    # 三个轴都归一化
    x_axis = normalize(x_axis)
    y_axis = normalize(y_axis)
    z_axis = normalize(z_axis)

    # 基本正交性检查
    xy = abs(dot(x_axis, y_axis))
    yz = abs(dot(y_axis, z_axis))
    zx = abs(dot(z_axis, x_axis))

    if max(xy, yz, zx) > 0.02:
        raise ValueError(
            "输入的 X+/Y+/Z+ 不是相互垂直的坐标轴。\n"
            "请检查三个方向向量。"
        )

    # 右手系检查：
    # X × Y 应该等于 Z
    cross_xy = normalize(cross(x_axis, y_axis))
    if dot(cross_xy, z_axis) < 0:
        raise ValueError(
            "输入的 X+/Y+/Z+ 不是右手坐标系。\n"
            "必须满足 X+ × Y+ = Z+。"
        )

    pose = Mat([
        [x_axis[0], y_axis[0], z_axis[0], 0],
        [x_axis[1], y_axis[1], z_axis[1], 0],
        [x_axis[2], y_axis[2], z_axis[2], 0],
        [0,         0,         0,         1]
    ])

    fanuc = Pose_2_Fanuc(pose)

    return (
        fanuc[3],
        fanuc[4],
        fanuc[5],
        pose
    )


def z_and_x_reference_to_rxyz(z_direction, x_reference):
    """
    已知 Z+ 方向，以及一个“X+参考方向”，
    自动构造完整右手坐标系。

    X+参考方向不要求本身严格垂直 Z+。
    程序会把它投影到垂直于 Z+ 的平面。
    """

    z_axis = normalize(z_direction)
    x_ref = normalize(x_reference)

    # X参考方向投影到垂直 Z+ 的平面
    x_axis = sub(
        x_ref,
        scale(z_axis, dot(x_ref, z_axis))
    )

    if vec_length(x_axis) < 1e-8:
        raise ValueError(
            "Z+ 与 X+参考方向平行或接近平行，"
            "无法确定滚转方向。"
        )

    x_axis = normalize(x_axis)

    # 右手系：X × Y = Z
    # 因此 Y = Z × X
    y_axis = normalize(cross(z_axis, x_axis))

    return axis_to_rxyz(x_axis, y_axis, z_axis)


def rotate_flange_z(pose, angle_deg):
    """绕法兰自身 Z+ 轴右手旋转；从 Z+ 端朝原点看，正角为逆时针。"""
    if not math.isfinite(angle_deg):
        raise ValueError("旋转角度必须是有限数字。")
    angle = math.radians(angle_deg)
    c, s = math.cos(angle), math.sin(angle)
    rotation = Mat([
        [c, -s, 0, 0],
        [s,  c, 0, 0],
        [0,  0, 1, 0],
        [0,  0, 0, 1]
    ])
    # 右乘表示绕局部轴旋转，而不是基座 Z 轴。
    rotated = pose * rotation
    values = Pose_2_Fanuc(rotated)
    return values[3], values[4], values[5], rotated


class DirectionToRxyzGUI:
    def __init__(self, root):
        self.root = root
        self.root.title("CR5 法兰坐标系 → RoboDK Rxyz")
        self.root.geometry("960x880")
        self.root.minsize(900, 800)

        self.mode = tk.StringVar(value="full")
        self.rotation_var = tk.StringVar(value="0")
        self.rotation_direction = tk.StringVar(value="顺时针")

        self.x_vars = [tk.StringVar() for _ in range(3)]
        self.y_vars = [tk.StringVar() for _ in range(3)]
        self.z_vars = [tk.StringVar() for _ in range(3)]

        self._build_ui()

        # 默认使用你目前讨论的方向。
        # 注意：这里给的是“法兰 Z+”，不是工具 Z-。
        self._set_axis(self.z_vars, 0, -1, 0)

        # 一组与 Z+=(0,-1,0) 配套的右手坐标系：
        # X+=(1,0,0)
        # Y+=(0,0,1)
        self._set_axis(self.x_vars, 1, 0, 0)
        self._set_axis(self.y_vars, 0, 0, 1)

        self.calculate()

    def _build_ui(self):
        ttk.Label(
            self.root,
            text="CR5 法兰坐标系 X+/Y+/Z+ → RoboDK Fanuc/Motoman Rxyz",
            font=("Microsoft YaHei UI", 16, "bold")
        ).pack(pady=(15, 5))

        ttk.Label(
            self.root,
            text=(
                "现在同时考虑红色 X+、绿色 Y+、蓝色 Z+。"
                "三根轴共同决定完整姿态。"
            ),
            font=("Microsoft YaHei UI", 10)
        ).pack(pady=(0, 12))

        # ====================================================
        # 模式选择
        # ====================================================
        mode_frame = ttk.LabelFrame(
            self.root,
            text="计算方式",
            padding=10
        )
        mode_frame.pack(fill="x", padx=18, pady=6)

        ttk.Radiobutton(
            mode_frame,
            text="完整坐标轴模式：输入 X+ / Y+ / Z+",
            variable=self.mode,
            value="full",
            command=self._update_mode
        ).pack(anchor="w")

        ttk.Radiobutton(
            mode_frame,
            text="方向 + 滚转参考模式：输入 Z+，再给一个 X+参考方向",
            variable=self.mode,
            value="zx",
            command=self._update_mode
        ).pack(anchor="w", pady=(5, 0))

        # ====================================================
        # 完整坐标轴输入
        # ====================================================
        self.full_frame = ttk.LabelFrame(
            self.root,
            text="1A. 法兰三个正方向（世界坐标）",
            padding=10
        )
        self.full_frame.pack(fill="x", padx=18, pady=6)

        self._build_axis_row(
            self.full_frame, "X+（红色）", self.x_vars, 0
        )
        self._build_axis_row(
            self.full_frame, "Y+（绿色）", self.y_vars, 1
        )
        self._build_axis_row(
            self.full_frame, "Z+（蓝色）", self.z_vars, 2
        )

        # ====================================================
        # Z+ + X参考输入
        # ====================================================
        self.zx_frame = ttk.LabelFrame(
            self.root,
            text="1B. Z+方向 + X+滚转参考",
            padding=10
        )

        self._build_axis_row(
            self.zx_frame, "Z+（蓝色）", self.z_vars, 0
        )
        self._build_axis_row(
            self.zx_frame, "X+参考（红色）", self.x_vars, 1
        )

        # ====================================================
        # 快速测试
        # ====================================================
        preset_frame = ttk.LabelFrame(
            self.root,
            text="快速测试",
            padding=10
        )
        preset_frame.pack(fill="x", padx=18, pady=6)

        ttk.Button(
            preset_frame,
            text="图中方向：Z+=(0,-1,0)",
            command=self.preset_current
        ).pack(side="left", padx=5)

        ttk.Button(
            preset_frame,
            text="Z+=+X",
            command=lambda: self.preset_z(1, 0, 0)
        ).pack(side="left", padx=5)

        ttk.Button(
            preset_frame,
            text="Z+=+Y",
            command=lambda: self.preset_z(0, 1, 0)
        ).pack(side="left", padx=5)

        ttk.Button(
            preset_frame,
            text="Z+=+Z",
            command=lambda: self.preset_z(0, 0, 1)
        ).pack(side="left", padx=5)

        rotation_frame = ttk.LabelFrame(
            self.root, text="末端追加旋转（绕法兰自身 Z 轴）", padding=10
        )
        rotation_frame.pack(fill="x", padx=18, pady=6)
        ttk.Label(rotation_frame, text="角度（度，非负）：").grid(row=0, column=0)
        ttk.Entry(rotation_frame, textvariable=self.rotation_var, width=12).grid(
            row=0, column=1, padx=8
        )
        ttk.Combobox(
            rotation_frame, textvariable=self.rotation_direction,
            values=("顺时针", "逆时针"), state="readonly", width=10
        ).grid(row=0, column=2, padx=8)
        ttk.Label(
            rotation_frame,
            text="观察方向：从法兰 Z+ 端朝原点看。每次均相对输入姿态计算，不累加。"
        ).grid(row=1, column=0, columnspan=3, sticky="w", pady=(8, 0))

        # ====================================================
        # 操作
        # ====================================================
        button_frame = ttk.Frame(self.root)
        button_frame.pack(pady=10)

        ttk.Button(
            button_frame,
            text="计算 Rxyz",
            command=self.calculate
        ).pack(side="left", padx=8)

        ttk.Button(
            button_frame,
            text="清空",
            command=self.clear
        ).pack(side="left", padx=8)

        # ====================================================
        # 结果
        # ====================================================
        result_frame = ttk.LabelFrame(
            self.root,
            text="2. 计算结果",
            padding=10
        )
        result_frame.pack(
            fill="both",
            expand=True,
            padx=18,
            pady=6
        )

        self.result_text = tk.Text(
            result_frame,
            font=("Consolas", 11),
            wrap="none"
        )
        self.result_text.pack(
            side="left",
            fill="both",
            expand=True
        )

        scrollbar = ttk.Scrollbar(
            result_frame,
            orient="vertical",
            command=self.result_text.yview
        )
        scrollbar.pack(side="right", fill="y")

        self.result_text.configure(
            yscrollcommand=scrollbar.set
        )

        ttk.Label(
            self.root,
            text=(
                "注意：仅一个 Z+ 方向不能唯一确定 Rxyz；"
                "必须再规定 X+/Y+ 的滚转方向。"
            ),
            font=("Microsoft YaHei UI", 9)
        ).pack(pady=(3, 12))

    def _build_axis_row(self, parent, title, vars_, row):
        ttk.Label(
            parent,
            text=title,
            width=18,
            font=("Microsoft YaHei UI", 10, "bold")
        ).grid(
            row=row,
            column=0,
            padx=(4, 10),
            pady=5,
            sticky="w"
        )

        for i, (axis_name, var) in enumerate(
            zip(["X", "Y", "Z"], vars_)
        ):
            ttk.Label(
                parent,
                text=axis_name
            ).grid(
                row=row,
                column=1 + i * 2,
                padx=(3, 4)
            )

            ttk.Entry(
                parent,
                textvariable=var,
                width=12,
                justify="center"
            ).grid(
                row=row,
                column=2 + i * 2,
                padx=(0, 12)
            )

    def _update_mode(self):
        if self.mode.get() == "full":
            self.zx_frame.pack_forget()
            self.full_frame.pack(
                fill="x",
                padx=18,
                pady=6,
                before=self._find_widget("快速测试")
            )
        else:
            self.full_frame.pack_forget()
            self.zx_frame.pack(
                fill="x",
                padx=18,
                pady=6,
                before=self._find_widget("快速测试")
            )

    def _find_widget(self, text):
        # 简单返回当前界面中的第一个 LabelFrame，
        # 这里只用于控制布局；找不到时返回 self
        for widget in self.root.winfo_children():
            if isinstance(widget, ttk.LabelFrame):
                if widget.cget("text") == text:
                    return widget
        return self.root

    def _set_axis(self, vars_, x, y, z):
        vars_[0].set(str(x))
        vars_[1].set(str(y))
        vars_[2].set(str(z))

    def preset_current(self):
        self._set_axis(self.z_vars, 0, -1, 0)
        self._set_axis(self.x_vars, 1, 0, 0)
        self._set_axis(self.y_vars, 0, 0, 1)
        self.mode.set("full")
        self._update_mode()
        self.calculate()

    def preset_z(self, x, y, z):
        self._set_axis(self.z_vars, x, y, z)

        # 根据 Z+ 自动寻找一个简单的 X+参考方向
        if abs(x) < 0.9:
            self._set_axis(self.x_vars, 1, 0, 0)
        else:
            self._set_axis(self.x_vars, 0, 1, 0)

        self.mode.set("zx")
        self._update_mode()
        self.calculate()

    def _read_vec(self, vars_, name):
        try:
            values = [
                float(var.get().strip())
                for var in vars_
            ]
        except (ValueError, AttributeError):
            raise ValueError(
                "%s 的三个分量必须全部是数字。" % name
            )

        if not all(math.isfinite(v) for v in values):
            raise ValueError(
                "%s 不能包含 NaN 或无穷值。" % name
            )

        return tuple(values)

    def calculate(self):
        try:
            if self.mode.get() == "full":
                x_axis = self._read_vec(self.x_vars, "X+")
                y_axis = self._read_vec(self.y_vars, "Y+")
                z_axis = self._read_vec(self.z_vars, "Z+")
                rx, ry, rz, pose = axis_to_rxyz(x_axis, y_axis, z_axis)
                mode_text = "完整坐标轴模式：直接使用输入的 X+/Y+/Z+"
            else:
                z_axis = self._read_vec(self.z_vars, "Z+")
                x_ref = self._read_vec(self.x_vars, "X+参考")
                rx, ry, rz, pose = z_and_x_reference_to_rxyz(z_axis, x_ref)
                x_axis = (pose[0,0], pose[1,0], pose[2,0])
                y_axis = (pose[0,1], pose[1,1], pose[2,1])
                z_axis = (pose[0,2], pose[1,2], pose[2,2])
                mode_text = "Z+ + X+参考模式：X+参考已投影到垂直 Z+ 的平面"

            # 处理旋转角度
            angle_deg = float(self.rotation_var.get().strip())
            if not math.isfinite(angle_deg) or angle_deg < 0:
                raise ValueError("旋转角度必须是非负有限数字。")
            signed_angle = -angle_deg if self.rotation_direction.get() == "顺时针" else angle_deg
            rx, ry, rz, pose = rotate_flange_z(pose, signed_angle)

            # 提取旋转后的轴向量
            x_axis = (pose[0,0], pose[1,0], pose[2,0])
            y_axis = (pose[0,1], pose[1,1], pose[2,1])
            z_axis = (pose[0,2], pose[1,2], pose[2,2])

            # ===== 新增：回填姿态到输入框，实现连续累加 =====
            self._set_axis(self.x_vars, x_axis[0], x_axis[1], x_axis[2])
            self._set_axis(self.y_vars, y_axis[0], y_axis[1], y_axis[2])
            self._set_axis(self.z_vars, z_axis[0], z_axis[1], z_axis[2])
            # 切换模式到“完整坐标轴模式”，以便显示三个轴
            self.mode.set("full")
            self._update_mode()
            # ===================================================

            mode_text += (
                "\n追加旋转：%s %.6f°（从 Z+ 端朝原点看）"
                "\n绕法兰局部 Z 轴，右手角度 = %+.6f°"
                % (self.rotation_direction.get(), angle_deg, signed_angle)
            )

            result = (
                "========================================\n"
                "CR5 法兰坐标系 → RoboDK Rxyz\n"
                "========================================\n\n"
                "【计算模式】\n"
                "%s\n\n"
                "【最终法兰坐标轴（世界坐标）】\n"
                "X+ = (%+.6f, %+.6f, %+.6f)\n"
                "Y+ = (%+.6f, %+.6f, %+.6f)\n"
                "Z+ = (%+.6f, %+.6f, %+.6f)\n\n"
                "【旋转矩阵 R】\n"
                "[ %+.6f  %+.6f  %+.6f ]\n"
                "[ %+.6f  %+.6f  %+.6f ]\n"
                "[ %+.6f  %+.6f  %+.6f ]\n\n"
                "【RoboDK Fanuc/Motoman】\n"
                "Rx = %+.6f deg\n"
                "Ry = %+.6f deg\n"
                "Rz = %+.6f deg\n\n"
                "【可直接用于 RoboDK 的位姿】\n"
                "[0, 0, 0, %.6f, %.6f, %.6f]\n\n"
                "【轴方向说明】\n"
                "红色箭头 = X+\n"
                "绿色箭头 = Y+\n"
                "蓝色箭头 = Z+\n\n"
                "注意：\n"
                "这里的 Z+ 就是你图片中确认的法兰蓝色箭头。\n"
                "因此不再对输入 Z+ 取反。\n"
                % (
                    mode_text,
                    x_axis[0], x_axis[1], x_axis[2],
                    y_axis[0], y_axis[1], y_axis[2],
                    z_axis[0], z_axis[1], z_axis[2],
                    pose[0,0], pose[0,1], pose[0,2],
                    pose[1,0], pose[1,1], pose[1,2],
                    pose[2,0], pose[2,1], pose[2,2],
                    rx, ry, rz,
                    rx, ry, rz
                )
            )

            self.result_text.delete("1.0", tk.END)
            self.result_text.insert("1.0", result)

        except Exception as e:
            messagebox.showerror("计算失败", "%s: %s" % (type(e).__name__, e))

    def clear(self):
        self.rotation_var.set("0")
        self.rotation_direction.set("顺时针")
        for var in (
            self.x_vars +
            self.y_vars +
            self.z_vars
        ):
            var.set("")

        self.result_text.delete("1.0", tk.END)


def main():
    root = tk.Tk()

    DirectionToRxyzGUI(root)

    root.mainloop()


if __name__ == "__main__":
    main()

--- Python program TCP仿真_升级前备份_20260909_173616 ---
# -*- coding: utf-8 -*-
"""
RoboDK 仿真：单点 + 连续运动（支持 TCP / 关节混合，含导入导出）
- 单点：指定 TCP -> IK 检查 -> MoveJ/MoveL
- 连续：逐点添加 TCP/关节 -> 检查可达性 -> 批量执行
姿态格式：Fanuc/Motoman
"""

from robodk.robolink import *
from robodk.robomath import *

import tkinter as tk
from tkinter import ttk, filedialog
import threading
import math
import json
import itertools

SIM_SPEED = 50.0
ALLOW_SIMULATION = True
MOVEJ_FALLBACK_MAX_DEVIATION_MM = 50.0  # MoveL失败后，MoveJ轨迹允许偏离TCP直线段的最大距离

RDK = Robolink()
robot = RDK.Item('', ITEM_TYPE_ROBOT)

if not robot.Valid():
    RDK.ShowMessage("未找到机械臂！", False)
    raise Exception("未找到机械臂")

# ============================================================
# Fanuc/Motoman 转换
# ============================================================
def fanuc_values_to_pose(x, y, z, rx, ry, rz):
    return Fanuc_2_Pose([x, y, z, rx, ry, rz])

def pose_to_fanuc_values(pose):
    return Pose_2_Fanuc(pose)

# ============================================================
# 全局变量（单点）
# ============================================================
target_pose = None
target_joints = None
simulation_running = False

# ============================================================
# 全局变量（连续运动）
# ============================================================
trajectory_records = []          # 存储 {'type':'TCP'/'JOINT', 'values':[...], 'target':pose, 'joints':[...]}
record_text = None
traj_entries = None
traj_type = None
traj_singular = None          # 当前输入 TCP 是否标记为末端特异点
traj_j6_direction = None      # 特异点 J6 转动方向：+180 / -180

# ============================================================
# GUI 构建
# ============================================================
root = tk.Tk()
root.title("RoboDK - 机械臂仿真控制（轨迹预检升级版）")
root.geometry("1200x750")
root.resizable(True, True)

# ---- Notebook ----
notebook = ttk.Notebook(root)
notebook.pack(fill=tk.BOTH, expand=True, padx=10, pady=5)

# ============================================================
# 选项卡 1：单点运动（保留原有功能）
# ============================================================
tab_single = ttk.Frame(notebook)
notebook.add(tab_single, text="单点运动")

input_frame = tk.LabelFrame(tab_single, text="目标 TCP（Fanuc/Motoman 格式）")
input_frame.pack(fill=tk.X, padx=10, pady=10)

names = ["X (mm)", "Y (mm)", "Z (mm)", "Rx (deg)", "Ry (deg)", "Rz (deg)"]
defaults = ["0.000", "-241.500", "1047.000", "-90.000", "0.000", "180.000"]
entries_single = []

for i in range(6):
    tk.Label(input_frame, text=names[i]).grid(row=0, column=i*2, padx=5, pady=10)
    e = tk.Entry(input_frame, width=12)
    e.insert(0, defaults[i])
    e.grid(row=0, column=i*2+1, padx=5, pady=10)
    entries_single.append(e)

status_var = tk.StringVar(value="请输入目标点，然后点击“检查目标点”")
tk.Label(tab_single, textvariable=status_var, font=("Microsoft YaHei", 12, "bold")).pack(pady=8)

# 按钮框架
btn_frame_single = tk.Frame(tab_single)
btn_frame_single.pack(fill=tk.X, padx=10, pady=5)

check_button = tk.Button(btn_frame_single, text="检查目标点", command=lambda: check_target(entries_single, status_var, simulate_button, log), width=18, font=("Microsoft YaHei", 10, "bold"))
check_button.pack(side=tk.LEFT, padx=5)

simulate_button = tk.Button(btn_frame_single, text="开始 MoveJ 仿真", command=lambda: start_simulation(entries_single, status_var, simulate_button, check_button, log), width=20, font=("Microsoft YaHei", 10, "bold"), state=tk.DISABLED)
simulate_button.pack(side=tk.LEFT, padx=5)

tk.Button(btn_frame_single, text="停止仿真", command=lambda: stop_simulation(status_var, simulate_button, check_button, log), width=14).pack(side=tk.LEFT, padx=5)
tk.Button(btn_frame_single, text="读取当前 TCP", command=lambda: read_current_tcp(log), width=16).pack(side=tk.LEFT, padx=5)
tk.Button(btn_frame_single, text="当前 TCP → 输入框", command=lambda: current_tcp_to_input(entries_single, log), width=18).pack(side=tk.LEFT, padx=5)

# ---- 日志（放在最下面）----
log_frame = tk.LabelFrame(tab_single, text="日志")
log_frame.pack(fill=tk.BOTH, expand=True, padx=10, pady=10)

text_output = tk.Text(log_frame, font=("Consolas", 10), wrap=tk.NONE)
text_output.pack(side=tk.LEFT, fill=tk.BOTH, expand=True)

scroll_y = ttk.Scrollbar(log_frame, orient=tk.VERTICAL, command=text_output.yview)
scroll_y.pack(side=tk.RIGHT, fill=tk.Y)
text_output.configure(yscrollcommand=scroll_y.set)

# ============================================================
# 选项卡 2：连续运动（含导入导出）
# ============================================================
tab_traj = ttk.Frame(notebook)
notebook.add(tab_traj, text="连续运动")

# ---- 输入区域 ----
frame_traj_input = tk.LabelFrame(tab_traj, text="连续运动点输入：每次输入 1 个 TCP 点或 1 组关节角度，点击“检查并加入”")
frame_traj_input.pack(fill=tk.X, padx=10, pady=10)

type_frame = tk.Frame(frame_traj_input)
type_frame.pack(fill=tk.X, padx=8, pady=5)

tk.Label(type_frame, text="点类型：").pack(side=tk.LEFT, padx=3)

traj_type = tk.StringVar(value="TCP")

def _update_traj_labels_and_defaults():
    """切换 TCP/关节时更新标签和默认值"""
    names = ["X", "Y", "Z", "Rx", "Ry", "Rz"] if traj_type.get() == "TCP" else ["J1", "J2", "J3", "J4", "J5", "J6"]
    defaults = ["0.000", "-241.500", "1047.000", "-90.000", "0.000", "180.000"] if traj_type.get() == "TCP" else ["0.000"]*6
    for i, e in enumerate(traj_entries):
        for widget in traj_value_frame.grid_slaves(row=0, column=i*2):
            widget.configure(text=names[i])
        e.delete(0, tk.END)
        e.insert(0, defaults[i])

tk.Radiobutton(type_frame, text="TCP（X,Y,Z,Rx,Ry,Rz）", variable=traj_type, value="TCP", command=_update_traj_labels_and_defaults).pack(side=tk.LEFT, padx=8)
tk.Radiobutton(type_frame, text="关节（J1~J6）", variable=traj_type, value="JOINT", command=_update_traj_labels_and_defaults).pack(side=tk.LEFT, padx=8)

# ---- 末端特异点设置 ----
singular_frame = tk.Frame(tab_traj)
singular_frame.pack(fill=tk.X, padx=10, pady=2)
traj_singular = tk.BooleanVar(value=False)
traj_j6_direction = tk.IntVar(value=180)
tk.Checkbutton(
    singular_frame,
    text="标记当前 TCP 为末端特异点（跳过 IK，J6 直接转 180°）",
    variable=traj_singular
).pack(side=tk.LEFT, padx=3)
tk.Label(singular_frame, text="J6优先方向（不可行时自动反向）：").pack(side=tk.LEFT, padx=(15, 2))
tk.Radiobutton(singular_frame, text="+180°", variable=traj_j6_direction, value=180).pack(side=tk.LEFT)
tk.Radiobutton(singular_frame, text="-180°", variable=traj_j6_direction, value=-180).pack(side=tk.LEFT)

movej_check_frame = tk.Frame(tab_traj)
movej_check_frame.pack(fill=tk.X, padx=10, pady=2)
tk.Label(movej_check_frame, text="MoveJ兜底轨迹最大允许偏离TCP直线：").pack(side=tk.LEFT, padx=3)
movej_deviation_var = tk.DoubleVar(value=MOVEJ_FALLBACK_MAX_DEVIATION_MM)
tk.Entry(movej_check_frame, textvariable=movej_deviation_var, width=8).pack(side=tk.LEFT, padx=3)
tk.Label(movej_check_frame, text="mm（MoveL失败后，先检查MoveJ轨迹；超限则拒绝MoveJ）", fg="#555555").pack(side=tk.LEFT, padx=3)

traj_value_frame = tk.Frame(frame_traj_input)
traj_value_frame.pack(fill=tk.X, padx=8, pady=5)

traj_entries = []
tcp_defaults = ["0.000", "-241.500", "1047.000", "-90.000", "0.000", "180.000"]
for i in range(6):
    tk.Label(traj_value_frame, text=["X","Y","Z","Rx","Ry","Rz"][i]).grid(row=0, column=i*2, padx=3, pady=8)
    e = tk.Entry(traj_value_frame, width=12)
    e.grid(row=0, column=i*2+1, padx=4, pady=8)
    e.insert(0, tcp_defaults[i])
    traj_entries.append(e)

# ---- 连续运动按钮 ----
btn_traj_input = tk.Frame(tab_traj)
btn_traj_input.pack(fill=tk.X, padx=10, pady=5)

tk.Button(btn_traj_input, text="检查并加入当前点", command=lambda: add_and_check_trajectory_point(traj_type, traj_entries, trajectory_records, record_text, log, traj_singular, traj_j6_direction), width=22, bg="#2196F3", fg="white", font=("Microsoft YaHei", 10, "bold")).pack(side=tk.LEFT, padx=3)
tk.Button(btn_traj_input, text="读取当前TCP并写入", command=lambda: read_current_tcp_to_traj(traj_type, traj_entries, log), width=20).pack(side=tk.LEFT, padx=3)
tk.Button(btn_traj_input, text="读取当前关节并写入", command=lambda: read_current_joints_to_traj(traj_type, traj_entries, log), width=20).pack(side=tk.LEFT, padx=3)
tk.Button(btn_traj_input, text="清空当前输入", command=lambda: clear_trajectory_input(traj_type, traj_entries, log), width=16).pack(side=tk.LEFT, padx=3)

tk.Label(tab_traj, text="普通 TCP 用 IK 判断可达并检查连续段；关节点只做角度规范化。标记为末端特异点的 TCP 跳过 IK，仅在执行时让 J6 转 ±180°，其后的普通 TCP 重新正常 IK。", fg="#555555").pack(anchor=tk.W, padx=15, pady=3)

# ---- 已添加点列表 ----
frame_record = tk.LabelFrame(tab_traj, text="已检查通过的连续运动点（按加入顺序执行，可混合 TCP / 关节点）")
frame_record.pack(fill=tk.BOTH, expand=True, padx=10, pady=8)

record_text = tk.Text(frame_record, font=("Consolas", 10), height=6)
record_text.pack(fill=tk.BOTH, expand=True, padx=5, pady=5)

# ---- 点管理按钮 ----
btn_record_frame = tk.Frame(tab_traj)
btn_record_frame.pack(fill=tk.X, padx=10, pady=4)

tk.Button(btn_record_frame, text="删除最后一点", command=lambda: delete_last_record(trajectory_records, record_text, log), width=15).pack(side=tk.LEFT, padx=3)
tk.Button(btn_record_frame, text="清空全部点", command=lambda: clear_records(trajectory_records, record_text, log), width=15).pack(side=tk.LEFT, padx=3)
tk.Button(btn_record_frame, text="执行整段连续运动", command=lambda: execute_recorded_trajectory(trajectory_records, log), width=24, font=("Microsoft YaHei", 10, "bold"), bg="#4CAF50", fg="white").pack(side=tk.LEFT, padx=3)

# ---------- 新增：导入导出按钮 ----------
tk.Button(btn_record_frame, text="导出轨迹", command=lambda: export_trajectory(trajectory_records, log), width=12).pack(side=tk.LEFT, padx=3)
tk.Button(btn_record_frame, text="导入轨迹", command=lambda: import_trajectory(trajectory_records, record_text, log), width=12).pack(side=tk.LEFT, padx=3)
# --------------------------------------

tk.Label(tab_traj, text="特异点保持J1～J5不变，直接MoveJ转动J6；整段检查±180°两方向，优先无需整圈回绕的方案。", fg="#555555").pack(anchor=tk.W, padx=15, pady=4)

traj_status_var = tk.StringVar(value="升级版：特异点J6自动选择±180°，优先避免整圈回绕。")
tk.Label(tab_traj, textvariable=traj_status_var, anchor=tk.W, wraplength=1100).pack(fill=tk.X, padx=15)
traj_log_frame = tk.LabelFrame(tab_traj, text="连续运动日志 / 停止原因")
traj_log_frame.pack(fill=tk.X, padx=10, pady=5)
traj_log_output = tk.Text(traj_log_frame, font=("Consolas", 10), height=5, wrap=tk.WORD)
traj_log_output.pack(side=tk.LEFT, fill=tk.X, expand=True)
traj_log_scroll = ttk.Scrollbar(traj_log_frame, command=traj_log_output.yview)
traj_log_scroll.pack(side=tk.RIGHT, fill=tk.Y)
traj_log_output.configure(yscrollcommand=traj_log_scroll.set)

# ============================================================
# 核心函数（单点）
# ============================================================
def log(text):
    print(text)
    try:
        text_output.insert(tk.END, str(text) + "\n")
        text_output.see(tk.END)
        traj_log_output.insert(tk.END, str(text) + "\n")
        traj_log_output.see(tk.END)
        if str(text).strip():
            traj_status_var.set(str(text))
        root.update_idletasks()
    except:
        pass

def set_status(text):
    status_var.set(text)

def get_input_values(entries):
    try:
        return [float(e.get()) for e in entries]
    except ValueError:
        log("✕ 输入错误：所有值必须为数字。")
        set_status("输入错误")
        return None

def check_target(entries, status_var, simulate_button, log):
    global target_pose, target_joints
    simulate_button.config(state=tk.DISABLED)
    target_pose = None
    target_joints = None

    values = get_input_values(entries)
    if values is None:
        return

    x, y, z, rx, ry, rz = values
    log("")
    log("============================================================")
    log("开始检查目标点")
    log("============================================================")
    log(f"目标 TCP：X={x:.3f} Y={y:.3f} Z={z:.3f} Rx={rx:.3f} Ry={ry:.3f} Rz={rz:.3f}")

    try:
        pose = fanuc_values_to_pose(x, y, z, rx, ry, rz)
        joints = robot.SolveIK(pose)
    except Exception as e:
        log(f"✕ IK 检查发生错误：{e}")
        set_status("IK 检查失败")
        return

    if joints is None:
        log("✕ SolveIK 返回 None")
        set_status("目标点不可达 ✕")
        return

    q = joints.list()
    if q is None or len(q) < 6:
        log(f"✕ IK 无效：SolveIK 未返回 6 个关节值，实际={q}")
        set_status("目标点 IK 不可用 ✕")
        return

    # IK -> FK 闭环校验
    try:
        fk_pose = robot.SolveFK(joints)
        fk = pose_to_fanuc_values(fk_pose)
        pos_err = ((fk[0]-x)**2 + (fk[1]-y)**2 + (fk[2]-z)**2) ** 0.5
        ang_err = math.degrees(pose_angle(invH(pose) * fk_pose))
        log("")
        log(f"[DEBUG] IK -> FK 验证：FK={fk}, 位置误差={pos_err:.6f} mm, 相对姿态误差={ang_err:.6f} deg")
        if pos_err > 0.5 or ang_err > 0.5:
            log("✕ IK/FK 闭环误差过大，拒绝执行。")
            set_status("IK/FK 验证失败 ✕")
            return
        log("✓ IK/FK 闭环验证通过")
    except Exception as e:
        log(f"✕ IK/FK 验证失败：{e}")
        set_status("IK/FK 验证失败 ✕")
        return

    target_pose = pose
    target_joints = joints

    log("")
    log("✓ 目标点 IK 可达")
    log("满足条件的一组关节角：")
    for i in range(6):
        log(f"J{i+1} = {q[i]:.3f} deg")

    actual = pose_to_fanuc_values(target_pose)
    log("")
    log("RoboDK 对应的 Fanuc/Motoman 姿态：")
    log(f"X={actual[0]:.3f} Y={actual[1]:.3f} Z={actual[2]:.3f} Rx={actual[3]:.3f} Ry={actual[4]:.3f} Rz={actual[5]:.3f}")
    log("")
    log("现在可以点击“开始 MoveJ 仿真”。")
    set_status("目标点可达 ✓，MoveJ 仿真已启用")
    simulate_button.config(state=tk.NORMAL)

def start_simulation(entries, status_var, simulate_button, check_button, log):
    global simulation_running
    if target_pose is None:
        log("✕ 尚未通过目标点检查。")
        return
    if not ALLOW_SIMULATION:
        log("当前禁止仿真运动。")
        return
    if simulation_running:
        log("仿真正在运行，请稍候。")
        return

    simulation_running = True
    simulate_button.config(state=tk.DISABLED)
    check_button.config(state=tk.DISABLED)

    def worker():
        global simulation_running
        try:
            log("")
            log("============================================================")
            log("开始 RoboDK 仿真")
            log("============================================================")
            robot.setSpeed(SIM_SPEED)
            log(f"速度：{SIM_SPEED:.1f} mm/s")
            if target_joints is not None:
                q = target_joints.list()
                log("正在运动到目标点（MoveJ，使用 IK 关节）...")
                log(f"J = {[round(float(v), 6) for v in q[:6]]}")
                robot.MoveJ(q[:6])
            else:
                log("✕ 没有有效 IK 关节，拒绝执行 MoveJ。")
                set_status("没有有效 IK，未执行")
                return
            log("")
            log("✓ 仿真完成")
            set_status("仿真完成 ✓")
        except Exception as e:
            log("")
            log(f"✕ 仿真失败：{type(e).__name__}: {e}")
            set_status("仿真失败")
        finally:
            simulation_running = False
            root.after(0, lambda: check_button.config(state=tk.NORMAL))
            root.after(0, lambda: simulate_button.config(state=tk.NORMAL))

    threading.Thread(target=worker, daemon=True).start()

def stop_simulation(status_var, simulate_button, check_button, log):
    global simulation_running
    try:
        robot.Stop()
        log("已发送停止命令。")
        set_status("仿真已停止")
    except Exception as e:
        log(f"停止失败：{e}")
    simulation_running = False
    simulate_button.config(state=tk.NORMAL)
    check_button.config(state=tk.NORMAL)

def read_current_tcp(log):
    try:
        pose = robot.Pose()
        values = pose_to_fanuc_values(pose)
        log("")
        log("============================================================")
        log("当前 RoboDK TCP（Fanuc/Motoman 格式）")
        log("============================================================")
        log(f"X={values[0]:.3f} Y={values[1]:.3f} Z={values[2]:.3f} Rx={values[3]:.3f} Ry={values[4]:.3f} Rz={values[5]:.3f}")
    except Exception as e:
        log(f"读取当前 TCP 失败：{e}")

def current_tcp_to_input(entries, log):
    try:
        pose = robot.Pose()
        values = pose_to_fanuc_values(pose)
        for e, val in zip(entries, values):
            e.delete(0, tk.END)
            e.insert(0, f"{val:.3f}")
        log("✓ 已将当前 RoboDK TCP 填入目标输入框。")
    except Exception as e:
        log(f"读取当前 TCP 失败：{e}")

# ============================================================
# 连续运动核心函数（移植自真实运动脚本，适配仿真）
# ============================================================

def refresh_record_list(record_text, trajectory_records):
    if record_text is None:
        return
    record_text.delete("1.0", tk.END)
    for i, rec in enumerate(trajectory_records, 1):
        kind = rec["type"]
        vals = rec["values"]
        if kind == "TCP":
            if rec.get("singular", False):
                sd = int(rec.get("j6_delta", 180))
                line = f"P{i:<3} [TCP-特异点 J6优先{sd:+d}°/可反向] X={vals[0]:9.3f} Y={vals[1]:9.3f} Z={vals[2]:9.3f} Rx={vals[3]:8.3f} Ry={vals[4]:8.3f} Rz={vals[5]:8.3f}\n"
            else:
                line = f"P{i:<3} [TCP]   X={vals[0]:9.3f} Y={vals[1]:9.3f} Z={vals[2]:9.3f} Rx={vals[3]:8.3f} Ry={vals[4]:8.3f} Rz={vals[5]:8.3f}\n"
        else:
            line = f"P{i:<3} [JNT]   J1={vals[0]:8.3f} J2={vals[1]:8.3f} J3={vals[2]:8.3f} J4={vals[3]:8.3f} J5={vals[4]:8.3f} J6={vals[5]:8.3f}\n"
        record_text.insert(tk.END, line)

def _parse_six_from_entries(entries, label):
    if not entries or len(entries) != 6:
        log(f"{label}输入框异常：需要 6 个值")
        return None
    try:
        vals = [float(e.get().strip()) for e in entries]
    except (ValueError, AttributeError):
        log(f"{label}输入无效：6 个值必须全部为数字")
        return None
    if not all(math.isfinite(v) for v in vals):
        log(f"{label}输入无效：不能包含 NaN 或无穷值")
        return None
    return vals

def _check_tcp_reachable(vals):
    """检查单个 TCP 点 IK 是否可达，返回 (True, target, joints)。"""
    try:
        target = fanuc_values_to_pose(*vals)
        joints = robot.SolveIK(target, tool=robot.PoseTool(), reference=robot.PoseFrame())
        if joints is None:
            log("TCP IK：不可达")
            return False, None, None
        q = joints.list()
        if len(q) < 6:
            log(f"TCP IK：返回关节数量异常：{q}")
            return False, None, None
        log("TCP IK：可达")
        log(f"  IK关节：J1={q[0]:.2f} J2={q[1]:.2f} J3={q[2]:.2f} J4={q[3]:.2f} J5={q[4]:.2f} J6={q[5]:.2f}")
        return True, target, q[:6]
    except Exception as e:
        log(f"TCP IK 检查失败：{type(e).__name__}: {e}")
        return False, None, None

def _check_tcp_segment_continuous(prev_vals, curr_vals, segment_index, samples=20):
    """检查相邻 TCP 点间插补路径的 IK 连续可达性"""
    if prev_vals is None:
        return True
    log(f"开始检查 P{segment_index-1} -> P{segment_index} 的 TCP 连续 IK（{samples+1} 个采样点）")
    for k in range(samples + 1):
        t = k / samples
        vals = [prev_vals[i] + (curr_vals[i] - prev_vals[i]) * t for i in range(6)]
        try:
            pose = fanuc_values_to_pose(*vals)
            joints = robot.SolveIK(pose)
            if joints is None:
                log(f"  P{segment_index-1} -> P{segment_index}：第 {k+1}/{samples+1} 个采样点 IK 不可达，t={t:.3f}")
                log(f"  TCP：X={vals[0]:.3f} Y={vals[1]:.3f} Z={vals[2]:.3f} Rx={vals[3]:.3f} Ry={vals[4]:.3f} Rz={vals[5]:.3f}")
                return False
            q = joints.list()
            if len(q) < 6:
                log(f"  P{segment_index-1} -> P{segment_index}：采样点 IK 返回异常：{q}")
                return False
        except Exception as e:
            log(f"  P{segment_index-1} -> P{segment_index}：采样点 IK 检查失败：{type(e).__name__}: {e}")
            return False
    log(f"P{segment_index-1} -> P{segment_index}：连续 IK 检查通过")
    return True

def add_and_check_trajectory_point(traj_type, traj_entries, trajectory_records, record_text, log, singular_var=None, j6_direction_var=None):
    kind = traj_type.get()
    vals = _parse_six_from_entries(traj_entries, kind)
    if vals is None:
        return

    log("")
    log(f"========== 检查连续运动第 {len(trajectory_records)+1} 点 ==========")

    # 末端特异点：用户明确声明该点只需要末端绕自身轴转 180°。
    # 因此完全跳过 SolveIK/连续 IK 检查，执行时只让 J6 转 ±180°。
    is_singular = bool(singular_var.get()) if singular_var is not None else False
    j6_delta = int(j6_direction_var.get()) if j6_direction_var is not None else 180

    if kind == "TCP" and is_singular:
        if not trajectory_records:
            log("末端特异点不能作为第一个点：需要先有一个起始运动点。")
            return
        if trajectory_records[-1]["type"] != "TCP" or trajectory_records[-1].get("singular", False):
            log("末端特异点前一项必须是普通 TCP 点；否则无法保证只是末端原地旋转 180°。")
            return
        prev_vals = trajectory_records[-1]["values"]
        pos_err = math.sqrt(sum((vals[k] - prev_vals[k]) ** 2 for k in range(3)))
        if pos_err > 1e-3:
            log("末端特异点未加入：它的 XYZ 必须与前一个普通 TCP 点相同。")
            log(f"  与前一点位置差：{pos_err:.6f} mm")
            log("  特异点的设计前提是：只改变末端绕自身轴的姿态，不改变 TCP 位置。")
            return
        try:
            target = fanuc_values_to_pose(*vals)
        except Exception as e:
            log(f"末端特异点姿态转换失败：{type(e).__name__}: {e}")
            return

        trajectory_records.append({
            "type": "TCP",
            "values": vals[:],
            "target": target,
            "joints": None,
            "singular": True,
            "j6_delta": j6_delta,
        })
        log(f"P{len(trajectory_records)} [TCP-特异点]：已加入，跳过 IK。")
        log(f"  执行时保持 J1~J5 不变，J6优先转 {j6_delta:+d}°；整段不可行时尝试反向。")
        log("  请确保该点与前一点相比确实只是末端绕自身轴旋转 180°。")
        refresh_record_list(record_text, trajectory_records)
        if singular_var is not None:
            singular_var.set(False)
        return

    if kind == "TCP":
        ok, target, joints = _check_tcp_reachable(vals)
        if not ok:
            log("该 TCP 点未加入轨迹。")
            return

        # 普通 TCP 与前一个普通 TCP 之间做连续 IK 检查。
        # 如果前一个点是末端特异点，则特异点本身跳过 IK；当前点从这里开始重新做普通 SolveIK，
        # 因此不把“特异点姿态 -> 当前姿态”当成普通 TCP 笛卡尔插补段。
        if trajectory_records and trajectory_records[-1]["type"] == "TCP" and not trajectory_records[-1].get("singular", False):
            prev_vals = trajectory_records[-1]["values"]
            segment_no = len(trajectory_records) + 1
            if not _check_tcp_segment_continuous(prev_vals, vals, segment_no, samples=20):
                log(f"P{segment_no} [TCP]：上一 TCP 点到当前 TCP 点的连续 IK 检查失败，该点未加入轨迹。")
                return

        trajectory_records.append({
            "type": "TCP",
            "values": vals[:],
            "target": target,
            "joints": joints,
        })
        log(f"P{len(trajectory_records)} [TCP]：检查通过，已加入连续运动。")
    else:
        # 关节点：角度规范到 (-180, 180]
        corrected = [((v + 180.0) % 360.0) - 180.0 for v in vals]
        corrected = [180.0 if v <= -180.0 else v for v in corrected]
        if corrected != vals:
            log("关节点角度已自动纠正到 (-180°, 180°]：")
            log("  原始：" + "  ".join(f"J{i+1}={vals[i]:+.3f}°" for i in range(6)))
            log("  修正：" + "  ".join(f"J{i+1}={corrected[i]:+.3f}°" for i in range(6)))
        trajectory_records.append({
            "type": "JOINT",
            "values": corrected[:],
            "target": None,
            "joints": corrected[:],
        })
        log(f"P{len(trajectory_records)} [JNT]：未做 IK 可达性检查，角度规范化后已加入连续运动。")

    refresh_record_list(record_text, trajectory_records)

def _write_values_to_traj_entries(values, label):
    if not traj_entries or len(traj_entries) != 6:
        log(f"连续运动输入框异常：无法写入当前{label}")
        return False
    for e, val in zip(traj_entries, values[:6]):
        e.delete(0, tk.END)
        e.insert(0, f"{val:.3f}")
    log(f"当前{label}已写入选项卡3输入框")
    return True

def read_current_tcp_to_traj(traj_type, traj_entries, log):
    try:
        pose = robot.Pose()
        vals = pose_to_fanuc_values(pose)
        log("========== 读取当前 TCP -> 连续运动输入框 ==========")
        log(f"X={vals[0]:+.3f} Y={vals[1]:+.3f} Z={vals[2]:+.3f} Rx={vals[3]:+.3f} Ry={vals[4]:+.3f} Rz={vals[5]:+.3f}")
        if traj_type.get() != "TCP":
            traj_type.set("TCP")
            _update_traj_labels_and_defaults()
        return _write_values_to_traj_entries(vals, "TCP")
    except Exception as e:
        log(f"读取当前 TCP 失败：{type(e).__name__}: {e}")
        return False

def read_current_joints_to_traj(traj_type, traj_entries, log):
    try:
        joints = robot.SimulatorJoints()
        q = list(joints) if hasattr(joints, "__iter__") else [joints]
        if len(q) < 6:
            log(f"读取当前关节失败：SimulatorJoints 返回 {q}")
            return False
        q = q[:6]
        log("========== 读取当前关节 -> 连续运动输入框 ==========")
        log(f"J1={q[0]:+.3f} J2={q[1]:+.3f} J3={q[2]:+.3f} J4={q[3]:+.3f} J5={q[4]:+.3f} J6={q[5]:+.3f}")
        if traj_type.get() != "JOINT":
            traj_type.set("JOINT")
            _update_traj_labels_and_defaults()
        return _write_values_to_traj_entries(q, "关节")
    except Exception as e:
        log(f"读取当前关节失败：{type(e).__name__}: {e}")
        return False

def clear_trajectory_input(traj_type, traj_entries, log):
    if not traj_entries:
        return
    for e in traj_entries:
        e.delete(0, tk.END)
    if traj_type.get() == "TCP":
        defaults = ["0.000", "-241.500", "1047.000", "-90.000", "0.000", "180.000"]
    else:
        defaults = ["0.000"] * 6
    for e, val in zip(traj_entries, defaults):
        e.insert(0, val)
    log("当前输入已清空（恢复默认值）")

def delete_last_record(trajectory_records, record_text, log):
    if trajectory_records:
        rec = trajectory_records.pop()
        refresh_record_list(record_text, trajectory_records)
        log(f"已删除最后一点：P{len(trajectory_records)+1} [{rec['type']}]")
    else:
        log("当前没有可删除的连续运动点")

def clear_records(trajectory_records, record_text, log):
    trajectory_records.clear()
    refresh_record_list(record_text, trajectory_records)
    log("连续运动点列表已清空")

# ============================================================
# 新增：导入导出函数
# ============================================================
def export_trajectory(trajectory_records, log):
    """导出轨迹到 JSON 文件"""
    if not trajectory_records:
        log("没有可导出的轨迹点。")
        return
    filepath = filedialog.asksaveasfilename(defaultextension=".json", filetypes=[("JSON files", "*.json"), ("All files", "*.*")])
    if not filepath:
        return
    try:
        # 只导出类型和数值，不保存 target/joints（执行时重新计算）
        export_data = [{"type": rec["type"], "values": rec["values"], "singular": bool(rec.get("singular", False)), "j6_delta": int(rec.get("j6_delta", 180))} for rec in trajectory_records]
        with open(filepath, 'w') as f:
            json.dump(export_data, f, indent=2)
        log(f"轨迹已导出到：{filepath}")
    except Exception as e:
        log(f"导出失败：{e}")

def import_trajectory(trajectory_records, record_text, log):
    """从 JSON 文件导入轨迹"""
    filepath = filedialog.askopenfilename(defaultextension=".json", filetypes=[("JSON files", "*.json"), ("All files", "*.*")])
    if not filepath:
        return
    try:
        with open(filepath, 'r') as f:
            data = json.load(f)
        if not isinstance(data, list):
            raise ValueError("文件内容不是列表格式")
        # 验证每个元素
        for item in data:
            if not isinstance(item, dict) or 'type' not in item or 'values' not in item:
                raise ValueError("每个点必须包含'type'和'values'字段")
            if item['type'] not in ('TCP', 'JOINT'):
                raise ValueError(f"不支持的type: {item['type']}")
            if not isinstance(item['values'], list) or len(item['values']) != 6:
                raise ValueError("values必须为长度为6的列表")
            for v in item['values']:
                if not isinstance(v, (int, float)):
                    raise ValueError(f"values中的值必须为数字: {v}")
        # 清空并加载（target/joints 置 None，执行时重新计算）
        trajectory_records.clear()
        for item in data:
            is_singular = bool(item.get("singular", False)) and item["type"] == "TCP"
            trajectory_records.append({
                "type": item["type"],
                "values": item["values"][:],
                "target": fanuc_values_to_pose(*item["values"]) if item["type"] == "TCP" else None,
                "joints": None,
                "singular": is_singular,
                "j6_delta": int(item.get("j6_delta", 180)) if is_singular else 0
            })
        refresh_record_list(record_text, trajectory_records)
        log(f"已从 {filepath} 导入 {len(data)} 个点")
    except Exception as e:
        log(f"导入失败：{e}")

# ============================================================
# MoveJ 兜底轨迹检查
# ============================================================
def _point_to_segment_distance(p, a, b):
    """3D点到线段距离，单位mm。"""
    ax, ay, az = a
    bx, by, bz = b
    px, py, pz = p
    ab = (bx-ax, by-ay, bz-az)
    ap = (px-ax, py-ay, pz-az)
    ab2 = ab[0]*ab[0] + ab[1]*ab[1] + ab[2]*ab[2]
    if ab2 < 1e-12:
        return math.sqrt((px-ax)**2 + (py-ay)**2 + (pz-az)**2)
    t = (ap[0]*ab[0] + ap[1]*ab[1] + ap[2]*ab[2]) / ab2
    t = max(0.0, min(1.0, t))
    q = (ax+t*ab[0], ay+t*ab[1], az+t*ab[2])
    return math.sqrt((px-q[0])**2 + (py-q[1])**2 + (pz-q[2])**2)


def _tcp_position_from_joints(q):
    """关节角 -> 当前参考坐标系下的TCP位置，与轨迹输入使用同一坐标系。"""
    f = pose_to_fanuc_values(invH(robot.PoseFrame()) * robot.SolveFK(q) * robot.PoseTool())
    return (float(f[0]), float(f[1]), float(f[2]))


def _check_movej_tcp_trajectory(start_q, target_q, start_tcp_vals, target_tcp_vals, log, samples=30, max_deviation_mm=None):
    """
    在真正执行MoveJ之前，用关节空间线性插补采样，计算TCP轨迹相对
    起点-终点TCP直线段的最大偏离距离。

    目的：MoveL失败时，不再无条件MoveJ；只有MoveJ造成的TCP空间绕行
    没有超过允许值，才允许用MoveJ兜底。
    """
    if max_deviation_mm is None:
        max_deviation_mm = MOVEJ_FALLBACK_MAX_DEVIATION_MM

    start_q = [float(v) for v in start_q[:6]]
    target_q = [float(v) for v in target_q[:6]]
    a = (float(start_tcp_vals[0]), float(start_tcp_vals[1]), float(start_tcp_vals[2]))
    b = (float(target_tcp_vals[0]), float(target_tcp_vals[1]), float(target_tcp_vals[2]))

    log("开始检查 MoveJ 兜底轨迹：%d 个采样点，允许最大TCP偏离 %.3f mm" % (samples + 1, max_deviation_mm))
    max_dev = -1.0
    max_info = None

    for k in range(samples + 1):
        t = float(k) / float(samples)
        q = [start_q[j] + (target_q[j] - start_q[j]) * t for j in range(6)]
        try:
            p = _tcp_position_from_joints(q)
        except Exception as e:
            log("  MoveJ轨迹检查失败：第 %d/%d 个采样点 FK失败：%s: %s" % (k+1, samples+1, type(e).__name__, e))
            return False

        dev = _point_to_segment_distance(p, a, b)
        if dev > max_dev:
            max_dev = dev
            max_info = (k, t, q, p)

        if dev > max_deviation_mm:
            log("✕ MoveJ兜底轨迹拒绝：第 %d/%d 个采样点偏离TCP直线 %.3f mm > %.3f mm" %
                (k+1, samples+1, dev, max_deviation_mm))
            log("  t=%.3f  TCP=(%.3f, %.3f, %.3f)" % (t, p[0], p[1], p[2]))
            log("  因此不会执行这个MoveJ兜底动作，避免出现不可接受的大绕圈。")
            return False

    if max_info is not None:
        k, t, q, p = max_info
        log("✓ MoveJ兜底轨迹检查通过")
        log("  最大TCP偏离直线：%.3f mm（采样 %d/%d，t=%.3f）" % (max_dev, k+1, samples+1, t))
        log("  最大偏离点TCP=(%.3f, %.3f, %.3f)" % (p[0], p[1], p[2]))
    return True


# ============================================================
# 执行连续运动（MoveL失败时先检查MoveJ轨迹）
# ============================================================
def _trajectory_pose(q):
    return invH(robot.PoseFrame()) * robot.SolveFK(q) * robot.PoseTool()


def _linear_path_endpoint(start, target):
    # 本机MoveL_Test返回成功后Joints()可能为全零；从插补矩阵读取实际终点。
    program = RDK.AddProgram('_TCP仿真_路径预检', robot)
    try:
        program.setVisible(False)
        robot.setJoints(start)
        program.setPoseFrame(robot.PoseFrame())
        program.setPoseTool(robot.PoseTool())
        program.MoveJ(start)
        program.MoveL(target)
        message, matrix, status = program.InstructionListJoints(mm_step=1, deg_step=1, collision_check=COLLISION_ON)
        if status < 0:
            return None, message
        end = matrix.tr().rows[-1][:6]
        error_pose = invH(target) * _trajectory_pose(end)
        if norm(error_pose.Pos()) > .01 or pose_angle(error_pose) > math.radians(.01):
            raise RuntimeError('路径预检返回的终点不匹配目标TCP。')
        return end, message
    finally:
        program.Delete()


def _trajectory_start_candidates(records, lower, upper):
    first_tcp = next((rec for rec in records if rec['type'] == 'TCP'), None)
    if first_tcp is None:
        return [None]
    pose = fanuc_values_to_pose(*first_tcp['values'])
    solutions = robot.SolveIK_All(pose, tool=robot.PoseTool(), reference=robot.PoseFrame())
    candidates = []
    for solution in solutions:
        q = [((float(v) + 180.0) % 360.0) - 180.0 for v in solution[:6]]
        if len(q) != 6:
            continue
        for turns6 in (0, -1, 1):
            candidate = q[:]
            candidate[5] += 360.0 * turns6
            if all(lower[j] <= candidate[j] <= upper[j] for j in range(6)):
                if not any(max(abs(a-b) for a, b in zip(candidate, old)) < 1e-6 for old in candidates):
                    candidates.append(candidate)
    # 与运行前的关节状态无关；先尝试靠近关节零位的解及其等效圈数。
    return sorted(candidates, key=lambda q: (sum(v*v for v in q), tuple(q)))


def _checked_j6_rewinds(q, lower, upper, max_deviation):
    """返回可实际执行的整圈回绕；TCP空间偏离和碰撞都必须通过检查。"""
    tcp = pose_to_fanuc_values(_trajectory_pose(q))
    for delta in (-360.0, 360.0):
        end = q[:]
        end[5] += delta
        if not lower[5] <= end[5] <= upper[5]:
            continue
        if not _check_movej_tcp_trajectory(q, end, tcp, tcp, lambda msg: None,
                                          samples=360, max_deviation_mm=max_deviation):
            continue
        if robot.MoveJ_Test(q, end, minstep_deg=1) == 0:
            yield end


def _plan_continuous_trajectory(records, max_deviation, log):
    if not math.isfinite(max_deviation) or max_deviation < 0:
        raise ValueError('MoveJ允许偏离必须是非负有限数。')
    for i, rec in enumerate(records):
        vals = rec['values']
        if rec['type'] not in ('TCP', 'JOINT') or len(vals) != 6 or not all(math.isfinite(v) for v in vals):
            raise ValueError(f'P{i+1}：点类型或六维数值无效。')
        if rec.get('singular', False):
            if rec['type'] != 'TCP' or i == 0 or records[i-1]['type'] != 'TCP' or records[i-1].get('singular', False):
                raise ValueError(f'P{i+1}：特异点必须紧跟普通TCP点。')
            if rec.get('j6_delta', 180) not in (-180, 180):
                raise ValueError(f'P{i+1}：J6方向必须为+180或-180。')
    saved = robot.Joints().list()[:6]
    lower, upper, _ = robot.JointLimits()
    lower, upper = lower.list(), upper.list()
    candidates = _trajectory_start_candidates(records, lower, upper)
    direction_choices = [(rec.get('j6_delta', 180), -rec.get('j6_delta', 180))
                         for rec in records if rec.get('singular', False)]
    last_error = '首个TCP没有限位内的逆解。'
    try:
        RDK.Render(False)
        # 先穷举特异点转向的整段组合；都不可行才允许额外整圈回绕。
        for allow_rewind, allow_fallback in ((False, False), (False, True), (True, False), (True, True)):
            failed_prefixes = set()
            for seed, directions in ((s, d) for s in candidates for d in itertools.product(*direction_choices)):
                seed_key = tuple(seed or [])
                if any((seed_key, directions[:n]) in failed_prefixes for n in range(len(directions)+1)):
                    continue
                selected_directions = iter(directions)
                direction_count = 0
                q = saved[:]
                first_tcp = True
                plan = []
                try:
                    for i, rec in enumerate(records, 1):
                        target = fanuc_values_to_pose(*rec['values']) if rec['type'] == 'TCP' else None
                        method, fallback = 'MoveJ', False
                        rewinds = []
                        selected_delta = None
                        special = rec.get('singular', False)
                        if rec['type'] == 'JOINT':
                            end = rec['values'][:]
                        elif special:
                            selected_delta = next(selected_directions)
                            direction_count += 1
                            end = q[:]
                            end[5] += selected_delta
                            if not lower[5] <= end[5] <= upper[5]:
                                if not allow_rewind:
                                    raise ValueError(f'P{i}：J6 {selected_delta:+d}°超限，尝试其他转向组合。')
                                for rewound in _checked_j6_rewinds(q, lower, upper, max_deviation):
                                    if lower[5] <= rewound[5] + selected_delta <= upper[5]:
                                        rewinds.append(rewound[:])
                                        q = rewound
                                        end = q[:]
                                        end[5] += selected_delta
                                        break
                                else:
                                    raise ValueError(f'P{i}：指定J6转向会超限，且没有通过偏离/碰撞检查的回绕。')
                            # 只改变J6，用FK核对目标位姿，不对特异点调用逆解。
                            error_pose = invH(target) * _trajectory_pose(end)
                            if norm(error_pose.Pos()) > 1e-3 or pose_angle(error_pose) > math.radians(.01):
                                raise ValueError(f'P{i}：仅旋转J6无法到达所标注TCP，请检查特异点标记/工具。')
                        elif first_tcp:
                            end = seed[:]
                            first_tcp = False
                        else:
                            end, detail = _linear_path_endpoint(q, target)
                            if end is None and allow_rewind:
                                for rewound in _checked_j6_rewinds(q, lower, upper, max_deviation):
                                    end, detail = _linear_path_endpoint(rewound, target)
                                    if end is not None:
                                        rewinds.append(rewound[:])
                                        q = rewound
                                        break
                            if end is not None:
                                method = 'MoveL'
                            else:
                                if not allow_fallback:
                                    raise ValueError(f'P{i}：MoveL路径检查失败：{detail}')
                                end = robot.SolveIK(target, q, robot.PoseTool(), robot.PoseFrame()).list()[:6]
                                if len(end) != 6 or not _check_movej_tcp_trajectory(q, end, pose_to_fanuc_values(_trajectory_pose(q)), rec['values'], lambda msg: None, samples=100, max_deviation_mm=max_deviation):
                                    raise ValueError(f'P{i}：MoveL不可行，MoveJ偏离超过{max_deviation:.3f} mm或无有效逆解。')
                                fallback = True
                        if not all(lower[j] <= end[j] <= upper[j] for j in range(6)):
                            raise ValueError(f'P{i}：关节超限，J6目标={end[5]:.3f}°。')
                        if method == 'MoveJ' and robot.MoveJ_Test(q, end, minstep_deg=1) != 0:
                            raise ValueError(f'P{i}：MoveJ路径检查失败。')
                        plan.append(dict(method=method, joints=end[:], special=special, fallback=fallback, rewinds=rewinds, j6_delta=selected_delta))
                        q = end[:]
                    log(f'整段路径预检通过：{len(plan)}点；首个TCP J6={seed[5]:+.3f}°。' if seed else f'整段路径预检通过：{len(plan)}个关节点。')
                    return plan
                except ValueError as exc:
                    # 后续尚未执行的J6方向不会改变已失败的路径前缀。
                    failed_prefixes.add((seed_key, directions[:direction_count]))
                    last_error = str(exc)
                    log(f'候选分支未通过：{last_error}')
        raise ValueError('没有找到整段可行的关节分支。' + last_error)
    finally:
        robot.setJoints(saved)
        RDK.Render(True)


def execute_recorded_trajectory(trajectory_records, log):
    global simulation_running
    if simulation_running:
        log('已有仿真正在运行，请等待结束。')
        return
    if not ALLOW_SIMULATION or not trajectory_records:
        log('当前禁止仿真或没有轨迹点。')
        return
    simulation_running = True
    completed_count = 0
    trace_owned = False
    i = 0
    try:
        RDK.setRunMode(RUNMODE_SIMULATE)
        if robot.Busy():
            raise RuntimeError('机器人正在执行其他动作，本次未启动。')
        trace_owned = True
        RDK.Command('Trace', 'Off')
        RDK.Command('Trace', 'Reset')
        records = [dict(rec, values=rec['values'][:]) for rec in trajectory_records]
        log(f'========== 整段路径预检：{len(records)}点（仿真模式） ==========')
        plan = _plan_continuous_trajectory(records, float(movej_deviation_var.get()), log)
        RDK.Command('Trace', 'Reset')
        RDK.Command('Trace', 'On')
        log('========== 正式仿真运动：现在仅显示本次实际运动轨迹 ==========')
        robot.setSpeed(SIM_SPEED)
        for i, step in enumerate(plan, 1):
            if RDK.RunMode() != RUNMODE_SIMULATE:
                raise RuntimeError('运行模式改变，停止仿真。')
            for rewound in step['rewinds']:
                before = robot.Joints().list()[:6]
                log(f'P{i}前：实际MoveJ回绕J6 {rewound[5]-before[5]:+.0f}°（{before[5]:+.3f}° → {rewound[5]:+.3f}°），已通过偏离及碰撞检查。')
                robot.MoveJ(rewound)
                if max(abs(a-b) for a, b in zip(robot.Joints().list()[:6], rewound)) > .1:
                    raise RuntimeError('回绕终点与预检关节不一致。')
            log(f'P{i} 开始 {step["method"]}，J6目标={step["joints"][5]:+.3f}°')
            # 执行预检得到的关节分支；运行时异常立即停止，不把停止/通信异常当作兜底请求。
            getattr(robot, step['method'])(step['joints'])
            actual = robot.Joints().list()[:6]
            if max(abs(a-b) for a, b in zip(actual, step['joints'])) > .1:
                raise RuntimeError('实际关节与预检终点不一致。')
            completed_count += 1
            suffix = f'（仅J6 {step["j6_delta"]:+d}°，J1～J5保持不变）' if step['special'] else ('（偏离检查后兜底）' if step['fallback'] else '')
            log(f'P{i} -> {step["method"]} 执行完成{suffix}')
        log(f'========== 连续运动仿真完成：{completed_count}/{len(plan)} 点 ==========')
    except Exception as exc:
        log(f'✕ 连续运动停止：已完成{completed_count}点，阶段={"路径预检" if i == 0 else "P"+str(i)}；{type(exc).__name__}: {exc}')
    finally:
        if trace_owned:
            RDK.Command('Trace', 'Off')
            RDK.Render(True)
        simulation_running = False


# ============================================================
# 启动信息
# ============================================================
log("程序准备完成。")
log(f"机器人：{robot.Name()}")
log("姿态格式：Fanuc/Motoman (XYZ mm, Rx/Ry/Rz deg)")
log("单点运动：输入 TCP -> 检查 IK -> 执行 MoveJ")
log("连续运动升级版：特异点直接关节MoveJ，仅J6自动选择±180°；优先整段无需回绕的方案，保留碰撞和偏离检查。")
log("新增：导入/导出轨迹（JSON 格式）")

root.mainloop()

